      def scale(value, rawRange, scaledRange):
          def computeSlope(inputRange, outputRange):
              outputRangeDelta = outputRange[1] - outputRange[0]
              inputRangeDelta = inputRange[1] - inputRange[0]

              if (inputRangeDelta == 0):
                  return 0
              else:
                  return outputRangeDelta / inputRangeDelta
              end
          end

          def computeIntercept(slope, inputRange, outputRange):
              return outputRange[0] - (slope * inputRange[0])
          end

          def clipScaledValue(outputScaledValue, outputRange):
              if (outputRange[0] < outputRange[1]):
                  return clipWhenLowerLimitIsLessThanHigher(outputScaledValue, outputRange)
              else:
                  return clipWhenLowerLimitIsGreaterThanHigherLimit(outputScaledValue, outputRange)
              end
          end

          def clipWhenLowerLimitIsGreaterThanHigherLimit(outputScaledValue, outputRange):
              if (outputScaledValue < outputRange[1]):
                  return outputRange[1]
              elif (outputScaledValue > outputRange[0]):
                  return outputRange[0]
              else:
                  return outputScaledValue
              end
          end

          def clipWhenLowerLimitIsLessThanHigher(outputScaledValue, outputRange):
              if (outputScaledValue < outputRange[0]):
                  return outputRange[0]
              elif (outputScaledValue > outputRange[1]):
                  return outputRange[1]
              else:
                  return outputScaledValue
              end
          end

          slope = computeSlope(rawRange, scaledRange)
          intercept = computeIntercept(slope, rawRange, scaledRange)
          scaledValue = slope * value + intercept
          return clipScaledValue(scaledValue, scaledRange)
      end

      def limit(value, range):
          return scale(value, range, range)
      end


  rq_init_comm_if_connected(9, "1")
  rq_init_comm_if_connected(2, "2")
  rq_init_comm_if_connected(3, "3")
  rq_init_comm_if_connected(4, "4")
  rq_print_connected_grippers()
  rq_gripper_communication_thread = run rq_gripper_communication()
  set_closed_norm(97.6470588235294, "1")
  set_open_norm(1.1764705882352942, "1")
  set_closed_mm(0.0, "1")
  set_open_mm(53.0, "1")
  set_closed_norm(100.0, "2")
  set_open_norm(0.0, "2")
  set_closed_mm(0.0, "2")
  set_open_mm(50.0, "2")
  set_closed_norm(100.0, "3")
  set_open_norm(0.0, "3")
  set_closed_mm(0.0, "3")
  set_open_mm(50.0, "3")
  set_closed_norm(100.0, "4")
  set_open_norm(0.0, "4")
  set_closed_mm(0.0, "4")
  set_open_mm(50.0, "4")
  rq_current_limit_enabled = False
  while(not rq_gripper_communication_thread_started):
      sleep(0.008)
  end
  # end: URCap Installation Node
  step_count_300fee78_b3e2_4ecc_acea_62356c60d52b = 0.0
  thread Step_Counter_Thread_351342f9_30f5_4523_8313_4ca12f4a91f7():
    while (True):
      step_count_300fee78_b3e2_4ecc_acea_62356c60d52b = step_count_300fee78_b3e2_4ecc_acea_62356c60d52b + 1.0
      sync()
    end
  end
  run Step_Counter_Thread_351342f9_30f5_4523_8313_4ca12f4a91f7()
  global AMR_Position=struct(position_identifier=0, x1=0, x2=0, y1=0, y2=0, theta1=0, theta2=0)
  global CAM_Pose=p[0,0,0,0,0,0]
  global CAM_Relation=""
  global CMD_Abort=  False
  global CMD_Clear=  False
  global CMD_Reset=  False
  global CMD_Start=  False
  global CMD_Suspend=  False
  global CMD_Unhold=  False
  global CMD_Unsuspend=  False
  global CNT_Rack_Output=0
  global FNC_Freedrive=  False
  global PRC_TubCounter=0
  global STP=0
  global easyPickCount_4=0
  global easyPickCount_7=0
  global easyPickNoObj_4=0
  global easyPickNoObj_7=0
  global easyPickParts_4=0
  global easyPickParts_7=0
  global TMR_Barcode=0
  global Container_mid_1_p=p[-.379239199143, -.127191311915, .299999999998, .000000000046, -.000000000021, -1.247199999994]
  global Container_mid_1_q=[-2.477408934449926, -1.2969853503591224, -1.875639182904262, -1.539621866126728, 1.5731943360401213, -2.8009955944022717]
  global trigger_otw_p=p[-.364831738276, -.163967193938, .343299997821, .000000000046, -.000000000020, -1.148401333327]
  global trigger_otw_q=[-2.378283213085033, -1.2994862387706814, -1.7634300687554951, -1.6493302004167063, 1.573123683454141, -2.8011223671816943]
  global Waypoint_54_p=p[.008800512419, -.547926542621, .402696567415, -.589884378425, -.007228654778, -.061268144704]
  global Waypoint_54_q=[-1.2044575850116175, -1.3416667741588135, -1.8272563219070435, -0.9884541195682068, 1.3621035814285278, -2.7712565104113978]
  global Waypoint_77_p=p[-.178371829612, -.433927395311, .368082383916, -.086593488055, .704679941724, -.007869906074]
  global Waypoint_77_q=[-1.265390698109762, -1.3355963987163086, -1.7944865226745605, -1.7402602634825648, 0.8780410885810852, -2.7713127771960657]
  global Waypoint_83_p=p[.008800512419, -.547926542621, .402696567415, -.589884378425, -.007228654778, -.061268144704]
  global Waypoint_83_q=[-1.2044575850116175, -1.3416667741588135, -1.8272563219070435, -0.9884541195682068, 1.3621035814285278, -2.7712565104113978]
  global Waypoint_84_p=p[-.178371829612, -.433927395311, .368082383916, -.086593488055, .704679941724, -.007869906074]
  global Waypoint_84_q=[-1.265390698109762, -1.3355963987163086, -1.7944865226745605, -1.7402602634825648, 0.8780410885810852, -2.7713127771960657]
  global Vial_above_1_p=p[.017105793010, -.652093028359, .184920586844, .000000000272, .000000000270, 1.564063451276]
  global Vial_above_1_q=[-1.3375440709712851, -1.9618096977868804, -1.4665759083780685, -1.2837941559171444, 1.5732503672317195, -4.47276330421513]
  global Vial_pick_poi_1_p=p[.017105792852, -.648922724010, .093307568731, .000000000271, .000000000270, 1.564063451276]
  global Vial_pick_poi_1_q=[-1.3366329456391917, -2.0375277831965413, -1.6071432798879028, -1.0675084332049813, 1.57309887265915, -4.471135348858068]
  global Waypoint_86_p=p[.019227646885, -.648669633640, .184920586950, .000000000000, .000000000000, .024063451426]
  global Waypoint_86_q=[-1.3331129109407733, -1.9540750545686123, -1.4775914902901128, -1.280581784992414, 1.5733500744865856, -2.928303704452631]
  global Waypoint_87_p=p[-.032361834699, -.348336136197, .391475576335, -.000008499254, .000014589902, -.004651426820]
  global Waypoint_87_q=[-1.2709335019096129, -1.1914598663441005, -1.708995335060501, -1.8117888533498316, 1.5729683532263925, -2.8379347397710237]
  global Vial_3FG_plac_1_p=p[-.031858676359, -.349402499566, .145301120695, .000000000000, .000000000000, .000000000000]
  global Vial_3FG_plac_1_q=[-1.2723975525801707, -1.252376585823825, -2.3128114007049496, -1.1470592278900167, 1.5730548099411423, -2.8414815174610535]
  global Waypoint_88_p=p[-.032361834699, -.348336136197, .391475576335, -.000008499254, .000014589902, -.004651426820]
  global Waypoint_88_q=[-1.2709335019096129, -1.1914598663441005, -1.708995335060501, -1.8117888533498316, 1.5729683532263925, -2.8379347397710237]
  global cap_dump_1_p=p[-.139168676487, -.420163541420, .146096395183, .000000000000, .000000000000, .000000000000]
  global cap_dump_1_q=[-1.584588644510994, -1.5093464179777323, -2.1118449369620347, -1.091059703602438, 1.5728943834877336, -3.154014906686923]
  global Waypoint_89_p=p[-.032361834699, -.348336136197, .391475576335, -.000008499254, .000014589902, -.004651426820]
  global Waypoint_89_q=[-1.2709335019096129, -1.1914598663441005, -1.708995335060501, -1.8117888533498316, 1.5729683532263925, -2.8379347397710237]
  global Vial_3FG_plac_2_p=p[-.031858676359, -.349402499566, .145301120695, .000000000000, .000000000000, .000000000000]
  global Vial_3FG_plac_2_q=[-1.2723975525801707, -1.252376585823825, -2.3128114007049496, -1.1470592278900167, 1.5730548099411423, -2.8414815174610535]
  global Waypoint_90_p=p[-.032361834699, -.348336136197, .391475576335, -.000008499254, .000014589902, -.004651426820]
  global Waypoint_90_q=[-1.2709335019096129, -1.1914598663441005, -1.708995335060501, -1.8117888533498316, 1.5729683532263925, -2.8379347397710237]
  global cap_dump_2_p=p[-.139168676487, -.420163541420, .146096395183, .000000000000, .000000000000, .000000000000]
  global cap_dump_2_q=[-1.584588644510994, -1.5093464179777323, -2.1118449369620347, -1.091059703602438, 1.5728943834877336, -3.154014906686923]
  global Waypoint_91_p=p[-.032361834699, -.348336136197, .391475576335, -.000008499254, .000014589902, -.004651426820]
  global Waypoint_91_q=[-1.2709335019096129, -1.1914598663441005, -1.708995335060501, -1.8117888533498316, 1.5729683532263925, -2.8379347397710237]
  global Vial_liq_abov_1_p=p[-.025303660977, -.338758622354, .426628485936, -1.315858642253, .800043520260, -.928295855026]
  global Vial_liq_abov_1_q=[-0.3789628187762659, -1.5149522957256814, -2.263045310974121, 0.7870649534412841, -0.750984017048971, -3.2237566153155726]
  global Vial_liq_pick_3_p=p[-.002660428945, -.335984893034, .159389832934, -1.150456778400, .673175527684, -1.010612657503]
  global Vial_liq_pick_3_q=[-0.3660772482501429, -1.4503649038127442, -2.4056053161621094, -1.994692941705221, 0.8039668202400208, -0.2508929411517542]
  global Vial_liq_pick_4_p=p[-.041402486291, -.356791603314, .125395323246, -1.143483969075, .651070210027, -.878721885453]
  global Vial_liq_pick_4_q=[-0.4426233705502476, -1.437252121513727, -2.551930962114307, -1.776528229806984, 0.6562026234073748, -0.43018811960029524]
  global Vial_liq_abov_2_p=p[-.025303660977, -.338758622354, .426628485936, -1.315858642253, .800043520260, -.928295855026]
  global Vial_liq_abov_2_q=[-0.3789628187762659, -1.5149522957256814, -2.263045310974121, 0.7870649534412841, -0.750984017048971, -3.2237566153155726]
  global Liquid_midway_1_p=p[.057575295009, -.583081747994, .306414980749, -1.351675548728, .120935756539, -.096908606303]
  global Liquid_midway_1_q=[-0.895174805318014, -1.7035466633238734, -2.380953073501587, 0.631549521083496, 0.7706599235534668, -2.9455552736865442]
  global shake_3_p=p[.057574880217, -.583085370269, .306422893466, -1.360996190983, -.155555042453, -.438136255921]
  global shake_3_q=[-0.8951800505267542, -1.7035466633238734, -2.380937099456787, 0.6315542894550782, 0.7706599235534669, -2.5394540616517496]
  global shake_4_p=p[.057581636113, -.583090570002, .306439684073, -1.308767904323, .368530312677, .214926493520]
  global shake_4_q=[-0.8951714674579065, -1.7035395107665003, -2.380906343460083, 0.6315504747578125, 0.7706480026245118, -3.3161255787892268]
  global drop_above_3_p=p[.268235025993, -.467784390499, .226219872376, -1.027832627524, -.430841408251, 1.004603115937]
  global drop_above_3_q=[-0.935645882283346, -1.6663371525206507, -2.4252893924713135, 0.41966931402172847, 1.8470635414123535, -3.4600217978106897]
  global drop_above_4_p=p[.219042229014, -.470775657081, .133754190740, -.313004595901, -.344395319364, 1.500564994056]
  global drop_above_4_q=[-1.0601594887284795, -1.70046459045642, -2.0799996233759863, -0.7243227230676759, 1.9429634314685202, -4.115129153870795]
  global liq_tran_3_p=p[.213067510942, -.469567035397, .100231043184, .251862243732, .217902579404, 1.592812335393]
  global liq_tran_3_q=[-0.7789645168037476, -1.822364827406652, -1.8643518410805573, -1.252158963840138, 1.3768134449520435, -3.9328333233290254]
  global drop_above_5_p=p[.219042229014, -.470775657081, .133754190740, -.313004595901, -.344395319364, 1.500564994056]
  global drop_above_5_q=[-1.0601594887284795, -1.70046459045642, -2.0799996233759863, -0.7243227230676759, 1.9429634314685202, -4.115129153870795]
  global Waypoint_92_p=p[.187119460405, -.493959476151, .133754190608, -.313004596540, -.344395317757, 1.500564993991]
  global Waypoint_92_q=[-1.1418328121400876, -1.7310553375189475, -2.033634768766424, -0.772026910513711, 1.958578934631971, -4.201588449364511]
  global liq_tran_4_p=p[.195957706507, -.493022614126, .100231042689, .160718757180, .109807038912, 1.525321508623]
  global liq_tran_4_q=[-0.881740380645474, -1.8244526267589851, -1.865100964490387, -1.1608866323693583, 1.4631433601076713, -3.973915130363038]
  global drop_above_6_p=p[.219042229014, -.470775657081, .133754190740, -.313004595901, -.344395319364, 1.500564994056]
  global drop_above_6_q=[-1.0601594887284795, -1.70046459045642, -2.0799996233759863, -0.7243227230676759, 1.9429634314685202, -4.115129153870795]
  global drop_above_7_p=p[.268235025993, -.467784390499, .226219872376, -1.027832627524, -.430841408251, 1.004603115937]
  global drop_above_7_q=[-0.935645882283346, -1.6663371525206507, -2.4252893924713135, 0.41966931402172847, 1.8470635414123535, -3.4600217978106897]
  global Liquid_midway_2_p=p[.057575295009, -.583081747994, .306414980749, -1.351675548728, .120935756539, -.096908606303]
  global Liquid_midway_2_q=[-0.895174805318014, -1.7035466633238734, -2.380953073501587, 0.631549521083496, 0.7706599235534668, -2.9455552736865442]
  global Vial_drop_abo_1_p=p[.000324902251, -.648569523142, .221894115667, -.873462921366, 1.165852672573, -1.482720593185]
  global Vial_drop_abo_1_q=[-1.0576906334721352, -2.393016994184633, -0.9236232851859159, -2.5729213042279273, 0.7903331288549689, -0.33286325848155585]
  global Vial_liq_drop_1_p=p[.001020867953, -.647659915585, .092915870838, -.834762611599, 1.081942994823, -1.540647900176]
  global Vial_liq_drop_1_q=[-1.0631954168193474, -2.4447642951220825, -1.128811017825127, -2.1983115491972294, 0.8130148661460634, -0.38984988696911316]
  global Vial_drop_abo_2_p=p[.000324902251, -.648569523142, .221894115667, -.873462921366, 1.165852672573, -1.482720593185]
  global Vial_drop_abo_2_q=[-1.0576906334721352, -2.393016994184633, -0.9236232851859159, -2.5729213042279273, 0.7903331288549689, -0.33286325848155585]
  global Spatula_otw_p=p[-.038472058237, -.263141484147, .425351216717, -.000441582511, -.000128175490, 3.034387645854]
  global Spatula_otw_q=[-1.1888947506684495, -1.0083288774886814, -1.7052227056065874, -1.9984805067363443, 1.5730180972985317, 0.48793409320312264]
  global pick_spat_L_abv_p=p[.239059466375, -.067212518441, .280720723617, .000017217488, -.000484427718, 3.106837214660]
  global pick_spat_L_abv_q=[0.292765616142962, -0.8565557553273315, -2.140199892763044, -1.715349495646084, 1.573623142106424, 1.8984976776985687]
  global spat_L_pick_p=p[.242468789885, -.067301915011, .193171208067, .000017217488, -.000484427718, 3.106837214657]
  global spat_L_pick_q=[0.2867414378807389, -0.8600077002089179, -2.3629148016312627, -1.4891831672860159, 1.5737695566221115, 1.8933890858591198]
  global spat_L_lift_p=p[.245402002494, -.067432373551, .289049296496, .000017217490, -.000484427724, 3.106837214657]
  global spat_L_lift_q=[0.2834351187564135, -0.8798320076811592, -2.1119436738532986, -1.7203314352121302, 1.573588313403067, 1.8891054681654005]
  global spat_L_side_p=p[.247133573905, -.017633681797, .289062935631, .000017217490, -.000484427724, 3.106837214657]
  global spat_L_side_q=[0.49719173575848863, -0.8582398211168538, -2.1182130454788215, -1.735610316654931, 1.5735817737572706, 2.1028402698705397]
  global spat_L_up_p=p[.247135508752, -.017665230822, .397130746165, .000017217490, -.000484427724, 3.106837214657]
  global spat_L_up_q=[0.49854946074076967, -0.9346239623559676, -1.808280269374471, -1.969158816463132, 1.5731020084036995, 2.1031742024348157]
  global spat_M_up_p=p[.245495561680, -.112112573515, .420343789747, .000026293989, -.000477463067, 3.067686800858]
  global spat_M_up_q=[0.09017908059107435, -1.0134242235449396, -1.71728844067247, -1.9814399845077446, 1.573013686840385, 1.733759055129931]
  global spat_M_pick_p=p[.244673518506, -.111985070134, .192299022723, .000026293990, -.000477463072, 3.067686800901]
  global spat_M_pick_q=[0.08834054082534859, -0.9272467647495475, -2.3438023910348154, -1.4411029496965373, 1.5736983399628084, 1.7342144371718433]
  global spat_S_Up_7_p=p[.252087445596, -.159242094834, .423281604617, .000026293954, -.000477463070, 3.067686800855]
  global spat_S_Up_7_q=[-0.09804692328730358, -1.0862987822056382, -1.6788706463996483, -1.9470242450550348, 1.5730147401359813, 1.5455107082823842]
  global spat_S_Pick_4_p=p[.245377020686, -.158668022535, .192285730279, .000026293985, -.000477463062, 3.067686800840]
  global spat_S_Pick_4_q=[-0.10087203759495189, -1.011188488703386, -2.311978084495874, -1.3890267520590838, 1.5735990551056096, 1.5450562970948172]
  global spat_S_Up_8_p=p[.252087445596, -.159242094834, .423281604617, .000026293954, -.000477463070, 3.067686800855]
  global spat_S_Up_8_q=[-0.09804692328730358, -1.0862987822056382, -1.6788706463996483, -1.9470242450550348, 1.5730147401359813, 1.5455107082823842]
  global spat_flatM_up_p=p[.229022666361, -.211442909333, .418634047126, .000026293953, -.000477463083, 3.067686800888]
  global spat_flatM_up_q=[-0.30183372580416545, -1.1157042924275036, -1.6775646144685776, -1.9189678841796578, 1.5730340557943228, 1.341766142011193]
  global spat_flatM_pick_p=p[.241028983327, -.208057297586, .192270533170, .000026293950, -.000477463079, 3.067686800885]
  global spat_flatM_pick_q=[-0.2805687960562633, -1.1003763929487214, -2.271431297337675, -1.3404236887924883, 1.5734924238720627, 1.3653813047742556]
  global spat_flatS_up_p=p[.237651953780, -.253943828614, .403961222825, .000026293950, -.000477463092, 3.067686800841]
  global spat_flatS_up_q=[-0.42363550926974103, -1.1939944599502539, -1.6745915127240307, -1.843675057902054, 1.5731001874678698, 1.220082820532415]
  global spat_flatS_pick_p=p[.241325662334, -.251726327528, .192256842740, .000026293947, -.000477463087, 3.067686800841]
  global spat_flatS_pick_q=[-0.4144907797170738, -1.1967447109013012, -2.21926362252748, -1.2962499335425761, 1.5733885098427622, 1.2314402238866728]
  global spat_S_pick_p=p[.238158866340, -.157926795425, .192632100345, .000026293989, -.000477463069, 3.067686800857]
  global spat_S_pick_q=[-0.10084756991493293, -0.9881392730064915, -2.3204232610157494, -1.403630829593915, 1.5736254260650586, 1.5450653591083503]
  global spat_S_up_p=p[.244260523725, -.164466690315, .417087579736, .000026293988, -.000477463072, 3.067686800857]
  global spat_S_up_q=[-0.12101499604198729, -1.0718307017854336, -1.7023391702814736, -1.938028805938881, 1.573044424728474, 1.5226045951991447]
  global Waypoint_7_p=p[-.472820924474, .292439826233, .207418370237, -.137787250486, 2.177332259632, -2.152029714756]
  global Waypoint_7_q=[-2.911134078210732, -1.90240864358569, -1.968768330510411, -2.500365101593811, 0.11427687110891149, 0.0958980389250167]
  global Waypoint_8_p=p[-.357612884176, -.251084817998, .212379799667, -.858181193174, 1.714832512191, -1.687547565568]
  global Waypoint_8_q=[-1.620834863369681, -1.8936194567376496, -1.9821394403832038, -2.4599791457905273, 0.6296693672615152, 0.07625365420707819]
  global Decapp_above_3_p=p[-.013480295948, -.359153355979, .266194408367, -.879653555922, 1.646336924805, -1.709111068605]
  global Decapp_above_3_q=[-0.9632157249872035, -2.0163405763031657, -1.5968194594157152, -2.6579215719847085, 1.251243398585566, 0.047906446502667066]
  global Decapp_place_3_p=p[-.013480295890, -.359153356055, .160907502384, -.879653554902, 1.646336919740, -1.709111066456]
  global Decapp_place_3_q=[-0.9633402410919709, -2.1541179572356635, -1.6937729380888573, -2.4232786481058053, 1.2517342187662468, 0.04818402956922263]
  global Decapp_above_4_p=p[-.013480295948, -.359153355979, .266194408367, -.879653555922, 1.646336924805, -1.709111068605]
  global Decapp_above_4_q=[-0.9632157249872035, -2.0163405763031657, -1.5968194594157152, -2.6579215719847085, 1.251243398585566, 0.047906446502667066]
  global Waypoint_78_p=p[-.051450028091, -.519555688329, .365718563414, -1.287302938145, 1.077637394477, -1.218524965834]
  global Waypoint_78_q=[-0.9214276262416012, -1.8899696965062578, -1.4939326452510562, -2.840015661555725, 0.5585157189668353, 0.033997638875617575]
  global Waypoint_10_p=p[-.330595116596, .282932669854, .220236276291, 1.304675539882, .014233792938, -1.753932442581]
  global Waypoint_10_q=[-3.189526379253601, -1.8418198435143305, -1.7138504750370807, -2.182789974066381, 1.0126080912871243, -2.4455984844694645]
  global Waypoint_9_p=p[-.538777454962, .370695704977, .175030018143, -.317104215445, 2.082346543003, -2.037631421082]
  global Waypoint_9_q=[-3.1158871966457857, -1.998548595120492, -1.941797010061462, -2.2703530575838844, -0.27573365931009164, -0.06926782177267654]
  global Powder_wayp1_p=p[-.472820924474, .292439826233, .207418370237, -.137787250486, 2.177332259632, -2.152029714756]
  global Powder_wayp1_q=[-2.911134078210732, -1.90240864358569, -1.968768330510411, -2.500365101593811, 0.11427687110891149, 0.0958980389250167]
  global Waypoint_2_p=p[-.357612884176, -.251084817998, .212379799667, -.858181193174, 1.714832512191, -1.687547565568]
  global Waypoint_2_q=[-1.620834863369681, -1.8936194567376496, -1.9821394403832038, -2.4599791457905273, 0.6296693672615152, 0.07625365420707819]
  global Postions_otw_p=p[-.010896578244, -.533368729951, .288851175116, -1.233738470894, 1.195331112012, -1.207314088469]
  global Postions_otw_q=[-0.898791023514228, -2.078490033037677, -1.4499891355755317, -2.7624416226992476, 0.6570218891920963, 0.02136606178275929]
  global cont_A_otw_p=p[.070238108556, -.655257851554, .184611566008, -1.090601381517, 1.404822685081, -1.413645380264]
  global cont_A_otw_q=[-0.990969136335913, -2.7123780097559784, -0.5772671651193146, -3.0005537851220403, 0.84719335943793, 0.020652463706785973]
  global cont_B_otw_p=p[.256012899886, -.515433666916, .157862612232, -1.209199576153, 1.209199576154, -1.209199576153]
  global cont_B_otw_q=[-0.6068713783523112, -2.5251567701153963, -1.0126698074772102, -2.742679391438185, 0.9631140738765777, -0.0042246938882417595]
  global cont_C_otw_p=p[.319495487998, -.362719410364, .163846736977, -1.233784872294, 1.195277203291, -1.207325031551]
  global cont_C_otw_q=[-0.3611889651645974, -2.404603865546651, -1.2341573845076566, -2.650535279811077, 1.1944844573128257, 0.01638086594640864]
  global Waypoint_1_p=p[-.352029261722, -.424157832422, .472326578019, -.000004407962, .000020663369, -1.529709227737]
  global Waypoint_1_q=[-2.017015745614491, -1.7423968528991196, -1.0053357238485425, -1.9644715035904907, 1.5727249689896, -2.060727852912713]
  global Waypoint_5_p=p[.219993437017, -.447144142811, .462350040687, .000006087494, .000031090075, .000022232405]
  global Waypoint_5_q=[-0.8406239476037944, -1.5982534362206806, -1.1934200873248484, -1.9205794898315975, 1.5727336676986443, -2.4135960466995314]
  global cont_B_safe_p=p[.256012900841, -.515433666823, .234963258529, -1.209199574203, 1.209199576702, -1.209199577238]
  global cont_B_safe_q=[-0.5984778117169087, -2.477204487479997, -0.8976875250023646, -2.905631546928806, 0.9709012567976698, -0.00424039942746024]
  global PosA_up_p=p[.028578953747, -.638006009765, .227275735849, -1.090660933958, 1.404791542934, -1.413645191233]
  global PosA_up_q=[-1.0254743496427432, -2.565176838504783, -0.7558042274983681, -2.9696064674274343, 0.8129191411995651, 0.021444818458024387]
  global PosA_pick_p=p[.026918718687, -.640084889741, .097901147521, -1.090660933959, 1.404791542934, -1.413645191233]
  global PosA_pick_q=[-1.028821435558534, -2.6899890636403807, -0.8526126047665157, -2.7478942693937167, 0.8103607002888742, 0.021326778146411485]
  global PosB_up_p=p[.239472634782, -.492481416782, .220767759213, -1.233738470883, 1.195331111998, -1.207314088469]
  global PosB_up_q=[-0.5800230603397054, -2.4076296700885997, -1.0699783327330836, -2.8116344407747427, 0.9750472858169287, 0.017627507888886562]
  global PosB_pick_p=p[.240630296955, -.494558620171, .096392895280, -1.233740573549, 1.195309876041, -1.207293779132]
  global PosB_pick_q=[-0.5816146260408139, -2.553273721769836, -1.1376320925804277, -2.5983292591462153, 0.9740936784345416, 0.017625262979849232]
  global PosC_up_p=p[.241566602786, -.359249123455, .230260583862, -1.233738470888, 1.195331111997, -1.207314088449]
  global PosC_up_q=[-0.39573787962534546, -2.2019009616581497, -1.4115270142506517, -2.675987785326166, 1.160180741930842, 0.01687917643039505]
  global PosC_pick_p=p[.240633854030, -.361553124916, .093979792658, -1.233738470878, 1.195331111997, -1.207314088469]
  global PosC_pick_q=[-0.39992427526118757, -2.386042391328985, -1.4894374567278712, -2.414022930893381, 1.1566786195951169, 0.01712017454263659]
  global Pow_decap_up_p=p[-.017556487132, -.367519866742, .275835445416, -.605635182849, 1.892518157522, -1.890848751165]
  global Pow_decap_up_q=[-1.1272088681128203, -2.1173924123331025, -1.4250048354055203, -2.7485980486387676, 1.4193896902217862, 0.023247957637719453]
  global pow_decap_place_p=p[-.020433194420, -.368310202914, .161281291611, -.605635182838, 1.892518157522, -1.890848751163]
  global pow_decap_place_q=[-1.132360890531647, -2.2521863255983092, -1.5302136899970318, -2.5086176644751683, 1.4149282844269635, 0.02347140074572661]
  global Decap_above_p=p[-.031863883354, -.349974838955, .288042264213, .000000000000, .000000000000, .000000000000]
  global Decap_above_q=[-1.271900116540503, -1.1670201114602632, -1.989291655468758, -1.5559360538518163, 1.573255119759632, -2.842476569674073]
  global Decapp_p=p[-.031864263150, -.349974612700, .230259377740, .000000000000, .000000000000, .000000000000]
  global Decapp_q=[-1.2723555431601419, -1.1810456878410935, -2.1291754890757737, -1.4020263844320349, 1.5732701843074919, -2.842325632263757]
  global Cap_above_p=p[-.224192409203, -.629599568633, .257274081142, .000015605575, -.000015166009, -1.647823825902]
  global Cap_above_q=[-1.710642681834492, -1.9674285251810462, -1.2705185053146897, -1.4742193161331247, 1.573506065067499, -1.6347709465008595]
  global Cap_place_p=p[-.224189049846, -.629597879697, .041885651757, .000015605572, -.000015166011, -1.647823825903]
  global Cap_place_q=[-1.7111696563854295, -2.13979870939016, -1.5941008764912503, -0.978265561728648, 1.5732789016410962, -1.6336328794662904]
  global OP_PowderA2_p=p[.009371277507, -.409434369247, .294169017766, -.823281033205, 1.709410851243, -1.698303593897]
  global OP_PowderA2_q=[-0.9994544761745754, -2.1395254572673217, -1.3437567783153916, -2.8143375616690456, 1.2617899549595724, 0.019614613715634555]
  global Decap_up_p=p[-.018339217391, -.367674469480, .249553854268, -.546164737599, 1.935964719000, -1.930057109666]
  global Decap_up_q=[-1.158124747223252, -2.1569920012936787, -1.4340832185069745, -2.7006032680036753, 1.4556626828962336, 0.02060977878679182]
  global Decap_pick_p=p[-.020429098827, -.367971872627, .161604333799, -.546164737600, 1.935964719000, -1.930057109666]
  global Decap_pick_q=[-1.161653098289774, -2.263509236689538, -1.5087211318402236, -2.519459740767391, 1.452646640403743, 0.02077912034002202]
  global Op_PowA_wP_p=p[-.173727579245, -.372934016396, .295116627479, -.972390492433, 1.540962074418, -1.548745344994]
  global Op_PowA_wP_q=[-1.1740587397768483, -1.865656321049359, -1.7426943793777419, -2.679427276872525, 0.8588908769087338, 0.017944699631825187]
  global TMR_Barcode_is_counting=False
  thread Timer_Thread():
    while (True):
      if (TMR_Barcode_is_counting):
        TMR_Barcode = TMR_Barcode + get_steptime()
      end
      sync()
    end
  end
  run Timer_Thread()
  def Sub_Vision_V18():
    $ 816 "Sub_Vision_V18" "noBreak"
    $ 817 "PreSettings"
    $ 818 "CAM_LM_Detected≔ False "
    global CAM_LM_Detected=  False
    $ 819 "CAM_Captures≔0"
    global CAM_Captures=0
    $ 820 "CAM_Pose≔p[0,0,0,0,0,0]"
    global CAM_Pose=p[0,0,0,0,0,0]
    $ 821 "CAM_LM_Refinmnt≔ False "
    global CAM_LM_Refinmnt=  False
    $ 822 "CAM_LM_Refined≔ False "
    global CAM_LM_Refined=  False
    $ 823 "CAM_LM_Deviatn≔p[0,0,0,0,0,0]"
    global CAM_LM_Deviatn=p[0,0,0,0,0,0]
    $ 824 "CAM_LM_ID≔0"
    global CAM_LM_ID=0
    $ 825 "CAM_Done≔ False "
    global CAM_Done=  False
    $ 826 "CAM_CNT_Obj≔0"
    global CAM_CNT_Obj=0
    $ 827 "CAM_Result = []"
    CAM_Result = []
    $ 828 "OBJ_Detected≔ False "
    global OBJ_Detected=  False
    $ 829 "FRM_Reference≔p[0,0,0,0,0,0]"
    global FRM_Reference=p[0,0,0,0,0,0]
    $ 830 "'=========='"
    # '=========='
    $ 831 "Switch Action"
    switch_1 = Action
    $ 832 "Case 13"
    if (13 == switch_1):
    elif (15 == switch_1):
      $ 950 "Case 15"
    elif (131 == switch_1):
      $ 996 "Case 131"
      $ 997 "Read (SensoPart)"
      $ 998 "Action_Info≔'search for landmark'"
      global Action_Info="search for landmark"
      $ 999 "CAM_LM≔CAM_LMs[4]"
      global CAM_LM=CAM_LMs[4]
      $ 1000 "CAM_Relation≔CAM_LM.capture_relation"
      global CAM_Relation=CAM_LM.capture_relation
      $ 1001 "go to capture pose"
      $ 1004 "If ITM_ID≟1 and JIG≟7"
      if (ITM_ID == 1  and  JIG == 7):
        $ 1005 "PSE_T≔uLM_Cap_SSRack"
        global PSE_T=uLM_Cap_SSRack
      else:
        $ 1006 "ElseIf ITM_ID≟5 and JIG≟7"
        if (ITM_ID == 5  and  JIG == 7):
          $ 1007 "PSE_T≔FRM_Cap_SSRack"
          global PSE_T=FRM_Cap_SSRack
        else:
          $ 1010 "ElseIf ITM_ID≟1 and JIG≟15"
          if (ITM_ID == 1 and JIG == 15):
            $ 1011 "MoveJ"
            $ 1012 "Container_mid_1" "breakAfter"
            movej(get_inverse_kin(Container_mid_1_p, qnear=Container_mid_1_q), a=1.3962634015954636, v=1.0471975511965976, r=0.05)
            $ 1014 "PSE_T≔FRM_Container_const"
            global PSE_T=p[-0.5003348223692186,0.35061804815168285,0.41579001388808423,-5.092943187272062E-5,1.0145185065363121E-4,-2.764319258713288]
          else:
            $ 1015 "ElseIf ITM_ID≟1 and JIG≟21"
            if (ITM_ID == 1 and JIG == 21):
              $ 1016 "PSE_T≔FRM_PoTS_const"
              global PSE_T=p[-0.5403054403210852,-0.10910773999775857,0.4828,3.058497512721046E-6,2.3454853329357316E-5,-2.208510541952706]
            else:
              $ 1017 "ElseIf ITM_ID≟1 and JIG≟17"
              if (ITM_ID == 1 and JIG == 17):
                $ 1018 "MoveJ"
                $ 1019 "trigger_otw" "breakAfter"
                movej(get_inverse_kin(trigger_otw_p, qnear=trigger_otw_q), a=1.3962634015954636, v=1.0471975511965976, r=0.05)
                $ 1023 "PSE_T≔FRM_weigh_scale_const"
                global PSE_T=p[-0.3804866881697204,0.025744252835212,0.4723487455232425,-1.0445769542396123E-4,-1.924788411074358E-5,-2.1691978730572363]
              end
            end
          end
        end
      end
      $ 1024 "do_transition(PSE_T, keep_rxry=False)"
      do_transition(PSE_T, keep_rxry=False)
      $ 1025 "Set"
      set_tcp(p[0.0,0.0,0.161,3.1415,0.0,0.0])
      $ 1026 "MoveJ"
      $ 1027 "PSE_T" "breakAfter"
      movej(PSE_T, a=1.3962634015954636, v=1.7453292519943295)
      $ 1028 "CAM_Pose≔get_actual_tcp_pose()"
      global CAM_Pose= get_actual_tcp_pose ()
      $ 1029 "Loop  not CAM_Done and  not ERROR.FLAG and  not CMD_Stop"
      while (  not  CAM_Done  and    not  ERROR.FLAG  and    not  CMD_Stop):
        $ 1030 "adjust capture pose"
        $ 1031 "If CAM_LM_Detected and CAM_LM_Refinmnt"
        if (CAM_LM_Detected  and  CAM_LM_Refinmnt):
          $ 1032 "PSE_T≔p[0,0,0.300,0,0,0]"
          global PSE_T=p[0,0,0.300,0,0,0]
          $ 1033 "CAM_Pose≔PSE_T"
          global CAM_Pose=PSE_T
          $ 1034 "If  not is_reachable(FRM_Reference,[PSE_T])"
          if (  not  is_reachable(FRM_Reference,[PSE_T])):
            $ 1035 "Error"
            $ 1036 "set_error(ERROR_POSE_NOT_REACHABLE)"
            set_error(ERROR_POSE_NOT_REACHABLE)
          end
          $ 1037 "If  not ERROR.FLAG"
          if (  not  ERROR.FLAG):
            $ 1038 "MoveJ"
            $ 1039 "PSE_T" "breakAfter"
            set_tcp(p[0.0,0.0,0.161,0.0,0.0,0.0])
            movej(pose_trans(FRM_Reference, PSE_T), a=0.8726646259971648, v=1.3962634015954636)
            $ 1040 "CAM_LM_Refined≔ True "
            global CAM_LM_Refined=  True
          end
        else:
          $ 1041 "ElseIf  not CAM_LM_Detected and CAM_Captures>0"
          if (  not  CAM_LM_Detected  and  CAM_Captures>0):
            $ 1042 "MoveL"
            $ 1043 "If FRM_Reference≟p[0,0,0,0,0,0]"
            if (FRM_Reference == p[0,0,0,0,0,0]):
              $ 1044 "PSE_T≔get_random_pose(pose_ref=CAM_Pose, mode='cubic', range_max=[0.150,0.150,0.015])"
              global PSE_T=get_random_pose(pose_ref=CAM_Pose, mode="cubic", range_max=[0.150,0.150,0.015])
            else:
              $ 1049 "Else" "noBreak"
              $ 1050 "PSE_T≔get_random_pose(pose_ref=CAM_Pose, mode='rotation', range_max=[10,10,0])"
              global PSE_T=get_random_pose(pose_ref=CAM_Pose, mode="rotation", range_max=[10,10,0])
              $ 1051 "CAM_LM_Refined≔ True "
              global CAM_LM_Refined=  True
            end
            $ 1052 "If get_inverse_kin_has_solution(pose_trans(FRM_Reference, PSE_T))"
            if (get_inverse_kin_has_solution( pose_trans (FRM_Reference, PSE_T))):
              $ 1053 "Comment"
              # Comment
              $ 1054 "PSE_T" "breakAfter"
              set_tcp(p[0.0,0.0,0.161,3.1415,0.0,0.0])
              movel(pose_trans(FRM_Reference, PSE_T), a=0.03, v=0.05)
            else:
              $ 1055 "Else" "noBreak"
              $ 1056 "'If random pose is out of reach, set the initial cam pose'"
              # 'If random pose is out of reach, set the initial cam pose'
              $ 1057 "PSE_T≔CAM_Pose"
              global PSE_T=CAM_Pose
            end
          end
        end
        $ 1058 "Wait: 2.0"
        sleep(2.0)
        $ 1059 "trigger"
        $ 1060 "If ITM_ID≟1 and JIG≟7"
        if (ITM_ID == 1  and  JIG == 7):
          # begin: URCap Program Node
          #   Source: SensoPart VISOR Robotic, 2.0.6, SensoPart Industriesensorik GmbH
          #   Type: VISOR Trigger
          $ 1061 "# 1 VISOR Trigger"
          visor_changeJob(1, "Landmark_INVITE_2", 6000)
          visor_trigger(1, 6000, "arm")
          # end: URCap Program Node
        else:
          $ 1062 "ElseIf ITM_ID≟5 and JIG≟7"
          if (ITM_ID == 5  and  JIG == 7):
            # begin: URCap Program Node
            #   Source: SensoPart VISOR Robotic, 2.0.6, SensoPart Industriesensorik GmbH
            #   Type: VISOR Trigger
            $ 1063 "# 1 VISOR Trigger"
            visor_changeJob(1, "Landmark_INVITE_2", 6000)
            visor_trigger(1, 6000, "arm")
            # end: URCap Program Node
          else:
            $ 1064 "ElseIf ITM_ID≟13 and JIG≟7"
            if (ITM_ID == 13  and  JIG == 7):
              # begin: URCap Program Node
              #   Source: SensoPart VISOR Robotic, 2.0.6, SensoPart Industriesensorik GmbH
              #   Type: VISOR Trigger
              $ 1065 "# 1 VISOR Trigger"
              visor_changeJob(1, "Landmark_INVITE_2", 6000)
              visor_trigger(1, 6000, "arm")
              # end: URCap Program Node
            else:
              $ 1066 "ElseIf ITM_ID≟1 and JIG≟15"
              if (ITM_ID == 1 and JIG == 15):
                # begin: URCap Program Node
                #   Source: SensoPart VISOR Robotic, 2.0.6, SensoPart Industriesensorik GmbH
                #   Type: VISOR Trigger
                $ 1067 "# 1 VISOR Trigger"
                visor_changeJob(1, "Aztec_no_dot_pick", 6000)
                visor_trigger(1, 6000, "arm")
                # end: URCap Program Node
              else:
                $ 1068 "ElseIf ITM_ID≟1 and JIG≟21"
                if (ITM_ID == 1 and JIG == 21):
                  # begin: URCap Program Node
                  #   Source: SensoPart VISOR Robotic, 2.0.6, SensoPart Industriesensorik GmbH
                  #   Type: VISOR Trigger
                  $ 1069 "# 1 VISOR Trigger"
                  visor_changeJob(1, "PoTS", 6000)
                  visor_trigger(1, 6000, "arm")
                  # end: URCap Program Node
                else:
                  $ 1070 "ElseIf ITM_ID≟1 and JIG≟17"
                  if (ITM_ID == 1 and JIG == 17):
                    # begin: URCap Program Node
                    #   Source: SensoPart VISOR Robotic, 2.0.6, SensoPart Industriesensorik GmbH
                    #   Type: VISOR Trigger
                    $ 1071 "# 1 VISOR Trigger"
                    visor_changeJob(1, "Weigh_target", 6000)
                    visor_trigger(1, 6000, "arm")
                    # end: URCap Program Node
                  end
                end
              end
            end
          end
        end
        $ 1075 "TM_3D_Found≔visor_partsFound(1)"
        global TM_3D_Found= visor_partsFound (1)
        $ 1077 "If TM_3D_Found>0"
        if (TM_3D_Found>0):
          $ 1078 "CAM_LM_Detected≔ True "
          global CAM_LM_Detected=  True
          $ 1079 "CAM_Captures≔0"
          global CAM_Captures=0
        else:
          $ 1080 "Else" "noBreak"
          $ 1081 "CAM_LM_Detected≔ False "
          global CAM_LM_Detected=  False
          $ 1082 "CAM_Captures≔CAM_Captures+1"
          global CAM_Captures=CAM_Captures+1
        end
        $ 1087 "result"
        $ 1088 "If CAM_LM_Detected"
        if (CAM_LM_Detected):
          $ 1089 "If (CAM_LM_Refinmnt and CAM_LM_Refined) or  not CAM_LM_Refinmnt"
          if ((CAM_LM_Refinmnt  and  CAM_LM_Refined)  or    not  CAM_LM_Refinmnt):
            $ 1147 "If ITM_ID≟1 and JIG≟7"
            if (ITM_ID == 1  and  JIG == 7):
              $ 1148 "CAM_LM_SSRack≔visor_getPose3d(1, 0)"
              global CAM_LM_SSRack= visor_getPose3d (1, 0)
            else:
              $ 1149 "ElseIf ITM_ID≟5 and JIG≟7"
              if (ITM_ID == 5  and  JIG == 7):
                $ 1150 "CAM_LM_SSRack≔visor_getPose3d(1, 0)"
                global CAM_LM_SSRack= visor_getPose3d (1, 0)
              else:
                $ 1153 "ElseIf ITM_ID≟1 and JIG≟15"
                if (ITM_ID == 1 and JIG == 15):
                  $ 1154 "CAM_LM_cont≔visor_getPose3d(1, 0)"
                  global CAM_LM_cont= visor_getPose3d (1, 0)
                  $ 1155 "Trigger≔get_actual_tcp_pose()"
                  global Trigger= get_actual_tcp_pose ()
                else:
                  $ 1156 "ElseIf ITM_ID≟1 and JIG≟21"
                  if (ITM_ID == 1 and JIG == 21):
                    $ 1157 "CAM_LM_cont≔visor_getPose3d(1, 0)"
                    global CAM_LM_cont= visor_getPose3d (1, 0)
                    $ 1158 "Trigger≔get_actual_tcp_pose()"
                    global Trigger= get_actual_tcp_pose ()
                  else:
                    $ 1159 "ElseIf ITM_ID≟1 and JIG≟17"
                    if (ITM_ID == 1 and JIG == 17):
                      $ 1160 "CAM_LM_cont≔visor_getPose3d(1, 0)"
                      global CAM_LM_cont= visor_getPose3d (1, 0)
                      $ 1161 "Trigger≔get_actual_tcp_pose()"
                      global Trigger= get_actual_tcp_pose ()
                    end
                  end
                end
              end
            end
            $ 1162 "CAM_Done≔ True "
            global CAM_Done=  True
          end
        else:
          $ 1163 "ElseIf  not CAM_LM_Detected and CAM_Captures<CAM_PRM_Retries"
          if (  not  CAM_LM_Detected  and  CAM_Captures<CAM_PRM_Retries):
            $ 1164 "CAM_LM_Refined≔ False "
            global CAM_LM_Refined=  False
          else:
            $ 1165 "ElseIf CAM_Captures≥CAM_PRM_Retries"
            if (CAM_Captures >= CAM_PRM_Retries):
              $ 1166 "CAM_Done≔ True "
              global CAM_Done=  True
              $ 1167 "Error"
              $ 1168 "set_error(ERROR_NO_LANDMARK)"
              set_error(ERROR_NO_LANDMARK)
            end
          end
        end
      end
    elif (151 == switch_1):
      $ 1169 "Case 151"
      $ 1170 "Detect (SensoPart)"
      $ 1171 "go to capture pose"
      $ 1172 "FRM_Reference≔FRM_Cap_SSRack"
      global FRM_Reference=FRM_Cap_SSRack
      $ 1173 "PSE_T≔p[0,0,-0.00,0,0,0]"
      global PSE_T=p[0,0,-0.00,0,0,0]
      $ 1174 "do_transition(pose_trans(FRM_Reference, PSE_T), keep_rxry=False)"
      do_transition( pose_trans (FRM_Reference, PSE_T), keep_rxry=False)
      $ 1175 "JNT_Q≔get_actual_joint_positions()"
      global JNT_Q= get_actual_joint_positions ()
      $ 1176 "JNT_Q≔[JNT_Q[0], JNT_Q[1], JNT_Q[2], JNT_Q[3], JNT_Q[4], 0]"
      global JNT_Q=[JNT_Q[0], JNT_Q[1], JNT_Q[2], JNT_Q[3], JNT_Q[4], 0]
      $ 1177 "Set"
      set_tcp(p[0.0,0.0,0.161,3.1415,0.0,0.0])
      $ 1178 "movej(get_inverse_kin(pose_trans(FRM_Reference, PSE_T), qnear=JNT_Q))"
      movej(get_inverse_kin( pose_trans (FRM_Reference, PSE_T), qnear=JNT_Q))
      $ 1179 "CAM_Pose≔pose_trans(pose_inv(FRM_Reference), get_actual_tcp_pose())"
      global CAM_Pose= pose_trans ( pose_inv (FRM_Reference),  get_actual_tcp_pose ())
      $ 1180 "Loop  not CAM_Done and  not ERROR.FLAG and  not CMD_Stop"
      while (  not  CAM_Done  and    not  ERROR.FLAG  and    not  CMD_Stop):
        $ 1181 "If  not OBJ_Detected and CAM_Captures>0"
        if (  not  OBJ_Detected  and  CAM_Captures>0):
          $ 1182 "MoveL"
          $ 1183 "If FRM_Reference≟p[0,0,0,0,0,0]"
          if (FRM_Reference == p[0,0,0,0,0,0]):
            $ 1185 "PSE_T≔get_random_pose(pose_ref=CAM_Pose, mode='rotation', range_max=[15,15,0])"
            global PSE_T=get_random_pose(pose_ref=CAM_Pose, mode="rotation", range_max=[15,15,0])
          else:
            $ 1186 "Else" "noBreak"
            $ 1187 "PSE_T≔get_random_pose(pose_ref=CAM_Pose, mode='rotation', range_max=[10,10,0])"
            global PSE_T=get_random_pose(pose_ref=CAM_Pose, mode="rotation", range_max=[10,10,0])
          end
          $ 1188 "If get_inverse_kin_has_solution(pose_trans(FRM_Reference, PSE_T))"
          if (get_inverse_kin_has_solution( pose_trans (FRM_Reference, PSE_T))):
            $ 1189 "PSE_T" "breakAfter"
            set_tcp(p[0.0,0.0,0.161,3.1415,0.0,0.0])
            movel(pose_trans(FRM_Reference, PSE_T), a=0.03, v=0.05)
          else:
            $ 1190 "Else" "noBreak"
            $ 1191 "'If random pose is out of reach, set the initial cam pose'"
            # 'If random pose is out of reach, set the initial cam pose'
            $ 1192 "PSE_T≔CAM_Pose"
            global PSE_T=CAM_Pose
            $ 1193 "PSE_T" "breakAfter"
            set_tcp(p[0.0,0.0,0.161,3.1415,0.0,0.0])
            movel(pose_trans(FRM_Reference, PSE_T), a=0.03, v=0.05)
          end
        end
        $ 1194 "Wait: 0.5"
        sleep(0.5)
        $ 1195 "Set"
        set_tcp(p[0.0,0.0,0.161,3.1415,0.0,0.0])
        # begin: URCap Program Node
        #   Source: SensoPart VISOR Robotic, 2.0.6, SensoPart Industriesensorik GmbH
        #   Type: VISOR Trigger
        $ 1196 "# 1 VISOR Trigger"
        visor_changeJob(1, "Object Detection Single", 6000)
        visor_trigger(1, 6000, "arm")
        # end: URCap Program Node
        $ 1197 "If visor_isResponseOk(1)"
        if ( visor_isResponseOk (1)):
          $ 1198 "CAM_CNT_Obj≔visor_partsFound(1)"
          global CAM_CNT_Obj= visor_partsFound (1)
          $ 1199 "CAM_OBJ_Pose≔visor_getPose3d(1, 0)"
          global CAM_OBJ_Pose= visor_getPose3d (1, 0)
          $ 1200 "If CAM_CNT_Obj>0"
          if (CAM_CNT_Obj>0):
            $ 1201 "CAM_OBJ_Color≔visor_getAdditionalData(1, 0)"
            global CAM_OBJ_Color= visor_getAdditionalData (1, 0)
            $ 1202 "CAM_DetectScore≔to_num(visor_getAdditionalData(1, 1))/1000"
            global CAM_DetectScore=to_num( visor_getAdditionalData (1, 1))/1000
            $ 1203 "OBJ_Detected≔ True "
            global OBJ_Detected=  True
          end
        else:
          $ 1204 "Else" "noBreak"
          $ 1205 "CAM_Captures≔CAM_Captures+1"
          global CAM_Captures=CAM_Captures+1
        end
        $ 1206 "If OBJ_Detected"
        if (OBJ_Detected):
          $ 1207 "Get object data"
          $ 1208 "PRC_CntDetect≔0"
          global PRC_CntDetect=0
          $ 1209 "Loop PRC_CntDetect<CAM_CNT_Obj"
          while (PRC_CntDetect<CAM_CNT_Obj):
            $ 1210 "get object and jig number"
            $ 1211 "If ITM_ID≟1 and JIG≟7"
            if (ITM_ID == 1  and  JIG == 7):
              $ 1212 "FRM_Reference≔FRM_Cap_SSRack"
              global FRM_Reference=FRM_Cap_SSRack
            else:
              $ 1213 "ElseIf ITM_ID≟5 and JIG≟7"
              if (ITM_ID == 5  and  JIG == 7):
                $ 1214 "FRM_Reference≔uLM_Cap_SSRack"
                global FRM_Reference=uLM_Cap_SSRack
              end
            end
            $ 1217 "PSE_T≔pose_trans(pose_inv(FRM_Reference), CAM_OBJ_Pose)"
            global PSE_T= pose_trans ( pose_inv (FRM_Reference), CAM_OBJ_Pose)
            $ 1218 "CAM_Result.append(get_pattern_counter(PSE_T, 'X', pattern=[10, 5], patternsize=[0.181, 0.081]))"
            CAM_Result.append(get_pattern_counter(PSE_T, "X", pattern=[10, 5], patternsize=[0.181, 0.081]))
            $ 1219 "PRC_CntDetect≔PRC_CntDetect+1"
            global PRC_CntDetect=PRC_CntDetect+1
          end
          $ 1220 "CAM_Done≔ True "
          global CAM_Done=  True
        else:
          $ 1221 "ElseIf CAM_Captures≥CAM_PRM_Retries"
          if (CAM_Captures >= CAM_PRM_Retries):
            $ 1222 "CAM_Done≔ True "
            global CAM_Done=  True
          else:
            $ 1223 "Else" "noBreak"
            $ 1224 "CAM_Captures≔CAM_Captures+1"
            global CAM_Captures=CAM_Captures+1
          end
        end
      end
    end
    $ 1225 "'=========='"
    # '=========='
    $ 1226 "PostSettings"
    $ 1227 "FRM_Reference≔p[0,0,0,0,0,0]"
    global FRM_Reference=p[0,0,0,0,0,0]
    $ 1228 "Set"
    set_tcp(p[0.0,0.0,0.161,3.1415,0.0,0.0])
    $ 1229 "CAM_Pose≔p[0,0,0,0,0,0]"
    global CAM_Pose=p[0,0,0,0,0,0]
    $ 1230 "Action≔0"
    global Action=0
    $ 1231 "Action_Info≔''"
    global Action_Info=""
  end
  def Sub_AMR_MiR_V3():
    $ 1232 "Sub_AMR_MiR_V3" "noBreak"
    $ 1233 "PreSettings"
    $ 1234 "AMR_TargetList≔[1,2,3,4,5,21,22,23,24,31,32,33,34,35,36,37,38,41]"
    global AMR_TargetList=[1,2,3,4,5,21,22,23,24,31,32,33,34,35,36,37,38,41]
    $ 1235 "AMR_Done≔ False "
    global AMR_Done=  False
    $ 1236 "AMR_PosActual≔T2O_Current_Pos"
    global AMR_PosActual=modbus_get_signal_status("T2O_Current_Pos")
    $ 1237 "AMR_Attemps≔T2O_Nav_Attemps"
    global AMR_Attemps=modbus_get_signal_status("T2O_Nav_Attemps")
    $ 1238 "AMR_Battery≔MiR_Battery_Lvl"
    global AMR_Battery=modbus_get_signal_status("MiR_Battery_Lvl")
    $ 1239 "AMR_Charging≔(T2O_Charging≟1)"
    global AMR_Charging=(modbus_get_signal_status("T2O_Charging") == 1)
    $ 1240 "AMR_Position≔struct(position_identifier=T2O_Current_Pos, x1=MiR_Position_X1, x2=MiR_Position_X2, y1=MiR_Position_Y1, y2=MiR_Position_Y2, theta1=MiR_Theta_1, theta2=MiR_Theta_2) "
    global AMR_Position=struct(position_identifier=modbus_get_signal_status("T2O_Current_Pos"), x1=modbus_get_signal_status("MiR_Position_X1"), x2=modbus_get_signal_status("MiR_Position_X2"), y1=modbus_get_signal_status("MiR_Position_Y1"), y2=modbus_get_signal_status("MiR_Position_Y2"), theta1=modbus_get_signal_status("MiR_Theta_1"), theta2=modbus_get_signal_status("MiR_Theta_2"))
    $ 1241 "If MiR_Mode≠7"
    if (modbus_get_signal_status("MiR_Mode") != 7):
      $ 1242 "Error"
      $ 1243 "set_error(ERROR_AMR_WRONG_MODE)"
      set_error(ERROR_AMR_WRONG_MODE)
      $ 1244 "AMR_Done≔ True "
      global AMR_Done=  True
    end
    $ 1245 "'=========='"
    # '=========='
    $ 1246 "Switch STATE"
    switch_1 = STATE
    $ 1247 "Case 1"
    if (1 == switch_1):
      $ 1248 "stopping"
      $ 1249 "If T2O_Done≟1 and O2T_Acknowledge≟0"
      if (modbus_get_signal_status("T2O_Done") == 1  and  modbus_get_signal_status("O2T_Acknowledge") == 0):
        $ 1250 "Set O2T_Acknowledge=1"
        modbus_set_output_register("O2T_Acknowledge", 1)
      end
      $ 1251 "Set MiR_CMD_Stop=On"
      modbus_set_output_signal("MiR_CMD_Stop", True)
      $ 1252 "AMR_Position.position_identifier = 0"
      AMR_Position.position_identifier = 0
      $ 1253 "AMR_Done≔ True "
      global AMR_Done=  True
    elif (2 == switch_1):
      $ 1254 "Case 2"
      $ 1255 "stopped"
      $ 1256 "If MiR_State≠3 and MiR_State≠5"
      if (modbus_get_signal_status("MiR_State") != 3  and  modbus_get_signal_status("MiR_State") != 5):
        $ 1257 "Set MiR_CMD_Stop=Off"
        modbus_set_output_signal("MiR_CMD_Stop", False)
      end
    elif (3 == switch_1):
      $ 1258 "Case 3"
      $ 1259 "resetting"
      $ 1260 "Set O2T_Mis_Main=Off"
      modbus_set_output_signal("O2T_Mis_Main", False)
      $ 1261 "Set O2T_Mis_Charge=Off"
      modbus_set_output_signal("O2T_Mis_Charge", False)
      $ 1262 "If MiR_Mis_Queue>0"
      if (modbus_get_signal_status("MiR_Mis_Queue")>0):
        $ 1263 "Set MiR_CMD_Clear_Q=On"
        modbus_set_output_signal("MiR_CMD_Clear_Q", True)
        $ 1264 "Wait MiR_Mis_Queue≟0"
        while (not(modbus_get_signal_status("MiR_Mis_Queue") == 0)):
          sync()
        end
        $ 1265 "Set MiR_CMD_Clear_Q=Off"
        modbus_set_output_signal("MiR_CMD_Clear_Q", False)
      end
      $ 1266 "If MiR_Error_ID≠0"
      if (modbus_get_signal_status("MiR_Error_ID") != 0):
        $ 1267 "Set MiR_CMD_Clear_E=On"
        modbus_set_output_signal("MiR_CMD_Clear_E", True)
        $ 1268 "Wait MiR_Error_ID≟0"
        while (not(modbus_get_signal_status("MiR_Error_ID") == 0)):
          sync()
        end
        $ 1269 "Set MiR_CMD_Clear_E=Off"
        modbus_set_output_signal("MiR_CMD_Clear_E", False)
      end
      $ 1270 "Set O2T_Action=0"
      modbus_set_output_register("O2T_Action", 0)
      $ 1271 "Set O2T_Acknowledge=0"
      modbus_set_output_register("O2T_Acknowledge", 0)
      $ 1272 "Set O2T_Target_Pos=0"
      modbus_set_output_register("O2T_Target_Pos", 0)
      $ 1273 "Set O2T_Footprint=0"
      modbus_set_output_register("O2T_Footprint", 0)
      $ 1274 "Set O2T_ProtectOff=0"
      modbus_set_output_register("O2T_ProtectOff", 0)
      $ 1275 "Set O2T_Dock=0"
      modbus_set_output_register("O2T_Dock", 0)
      $ 1276 "AMR_Attemps≔0"
      global AMR_Attemps=0
      $ 1277 "AMR_PosTarget≔0"
      global AMR_PosTarget=0
      $ 1278 "AMR_Step≔0"
      global AMR_Step=0
      $ 1279 "AMR_AtTarget≔ False "
      global AMR_AtTarget=  False
      $ 1280 "If MiR_State≟4 or MiR_State≟3 or MiR_State≟10"
      if (modbus_get_signal_status("MiR_State") == 4  or  modbus_get_signal_status("MiR_State") == 3  or  modbus_get_signal_status("MiR_State") == 10):
        $ 1281 "AMR_Done≔ True "
        global AMR_Done=  True
      end
    elif (5 == switch_1):
      $ 1282 "Case 5"
      $ 1283 "starting"
      $ 1284 "If MiR_State≟4"
      if (modbus_get_signal_status("MiR_State") == 4):
        $ 1285 "Set MiR_CMD_Start=On"
        modbus_set_output_signal("MiR_CMD_Start", True)
        $ 1286 "Wait MiR_State≠4"
        while (not(modbus_get_signal_status("MiR_State") != 4)):
          sync()
        end
        $ 1287 "Set MiR_CMD_Start=Off"
        modbus_set_output_signal("MiR_CMD_Start", False)
        $ 1288 "AMR_Done≔ True "
        global AMR_Done=  True
      else:
        $ 1289 "ElseIf MiR_State≟10"
        if (modbus_get_signal_status("MiR_State") == 10):
          $ 1290 "'MiR in protective stop. Wait'"
          # 'MiR in protective stop. Wait'
          $ 1291 "AMR_Done≔ True "
          global AMR_Done=  True
        else:
          $ 1292 "ElseIf MiR_State≟3"
          if (modbus_get_signal_status("MiR_State") == 3):
            $ 1293 "AMR_Done≔ True "
            global AMR_Done=  True
          end
        end
      end
    elif (6 == switch_1):
      $ 1294 "Case 6"
      $ 1295 "execute"
      $ 1296 "AMR_AtTarget≔(AMR_PosActual≟AMR_PosTarget)"
      global AMR_AtTarget=(AMR_PosActual == AMR_PosTarget)
      $ 1297 "Switch AMR_Step"
      switch_2 = AMR_Step
      $ 1298 "Case 0"
      if (0 == switch_2):
        $ 1299 "If  not AMR_AtTarget"
        if (  not  AMR_AtTarget):
          $ 1300 "AMR_Step≔1"
          global AMR_Step=1
        else:
          $ 1301 "Else" "noBreak"
          $ 1302 "AMR_Done≔ True "
          global AMR_Done=  True
        end
      elif (1 == switch_2):
        $ 1303 "Case 1"
        $ 1304 "general Settings"
        $ 1305 "Set O2T_Acknowledge=0"
        modbus_set_output_register("O2T_Acknowledge", 0)
        $ 1306 "check for error"
        $ 1307 "If OBJ_Picked and MiR_State≟10"
        if (OBJ_Picked  and  modbus_get_signal_status("MiR_State") == 10):
          $ 1308 "Error"
          $ 1309 "set_error(ERROR_ROBOT_ARM_NOT_IN_HOME_POSE)"
          set_error(ERROR_ROBOT_ARM_NOT_IN_HOME_POSE)
          $ 1310 "Action≔0"
          global Action=0
        else:
          $ 1311 "ElseIf  not found_in_list(AMR_PosTarget, AMR_TargetList)"
          if (  not  found_in_list(AMR_PosTarget, AMR_TargetList)):
            $ 1312 "Error"
            $ 1313 "set_error(ERROR_UNKNOWN_POSE)"
            set_error(ERROR_UNKNOWN_POSE)
            $ 1314 "Action≔0"
            global Action=0
          end
        end
        $ 1315 "If MiR_State≟3"
        if (modbus_get_signal_status("MiR_State") == 3):
          $ 1316 "Set MiR_CMD_Start=Off"
          modbus_set_output_signal("MiR_CMD_Start", False)
          $ 1317 "Switch Action"
          switch_3 = Action
          $ 1318 "Case 51"
          if (51 == switch_3):
            $ 1319 "Charge"
            $ 1320 "'trigger the charging mission'"
            # 'trigger the charging mission'
            $ 1321 "'target pos is predefined'"
            # 'target pos is predefined'
            $ 1322 "Set O2T_Footprint=0"
            modbus_set_output_register("O2T_Footprint", 0)
            $ 1323 "Set O2T_Action=1"
            modbus_set_output_register("O2T_Action", 1)
            $ 1324 "If MiR_Mis_Queue≟0"
            if (modbus_get_signal_status("MiR_Mis_Queue") == 0):
              $ 1325 "Set O2T_Mis_Charge=On"
              modbus_set_output_signal("O2T_Mis_Charge", True)
              $ 1326 "Wait MiR_Mis_Queue≥1"
              while (not(modbus_get_signal_status("MiR_Mis_Queue") >= 1)):
                sync()
              end
              $ 1327 "Set O2T_Mis_Charge=Off"
              modbus_set_output_signal("O2T_Mis_Charge", False)
            end
          elif (52 == switch_3):
            $ 1328 "Case 52"
            $ 1329 "Navigate"
            $ 1330 "'trigger the standard missoin'"
            # 'trigger the standard missoin'
            $ 1331 "Set O2T_Footprint=AMR_FootprintID"
            modbus_set_output_register("O2T_Footprint", AMR_FootprintID)
            $ 1332 "Set O2T_Target_Pos=AMR_PosTarget"
            modbus_set_output_register("O2T_Target_Pos", AMR_PosTarget)
            $ 1333 "Set O2T_Action=2"
            modbus_set_output_register("O2T_Action", 2)
            $ 1334 "If MiR_Mis_Queue≟0"
            if (modbus_get_signal_status("MiR_Mis_Queue") == 0):
              $ 1335 "Set O2T_Mis_Main=On"
              modbus_set_output_signal("O2T_Mis_Main", True)
              $ 1336 "Wait MiR_Mis_Queue≥1"
              while (not(modbus_get_signal_status("MiR_Mis_Queue") >= 1)):
                sync()
              end
              $ 1337 "Set O2T_Mis_Main=Off"
              modbus_set_output_signal("O2T_Mis_Main", False)
            end
          end
        else:
          $ 1338 "ElseIf MiR_State≟4"
          if (modbus_get_signal_status("MiR_State") == 4):
            $ 1339 "Set MiR_CMD_Start=On"
            modbus_set_output_signal("MiR_CMD_Start", True)
          else:
            $ 1340 "ElseIf MiR_State≟5"
            if (modbus_get_signal_status("MiR_State") == 5):
              $ 1341 "AMR_Step≔2"
              global AMR_Step=2
            else:
              $ 1342 "ElseIf MiR_State≟10"
              if (modbus_get_signal_status("MiR_State") == 10):
                $ 1343 "'AMR still in safeguard stop'"
                # 'AMR still in safeguard stop'
              end
            end
          end
        end
      elif (2 == switch_2):
        $ 1344 "Case 2"
        $ 1345 "acknowledge handshake"
        $ 1346 "If T2O_Done≟1 and O2T_Acknowledge≟0"
        if (modbus_get_signal_status("T2O_Done") == 1  and  modbus_get_signal_status("O2T_Acknowledge") == 0):
          $ 1347 "Set O2T_Acknowledge=1"
          modbus_set_output_register("O2T_Acknowledge", 1)
        else:
          $ 1348 "ElseIf T2O_Done≟0 and O2T_Acknowledge≟1"
          if (modbus_get_signal_status("T2O_Done") == 0  and  modbus_get_signal_status("O2T_Acknowledge") == 1):
            $ 1349 "Set O2T_Acknowledge=0"
            modbus_set_output_register("O2T_Acknowledge", 0)
            $ 1350 "AMR_AtTarget≔(AMR_PosActual≟AMR_PosTarget)"
            global AMR_AtTarget=(AMR_PosActual == AMR_PosTarget)
            $ 1351 "AMR_Done≔ True "
            global AMR_Done=  True
          end
        end
      end
      $ 1352 "translate errors"
      $ 1353 "If AMR_Done"
      if (AMR_Done):
        $ 1354 "Switch T2O_Error_ID"
        switch_2 = modbus_get_signal_status("T2O_Error_ID")
        $ 1355 "Case 2003"
        if (2003 == switch_2):
          $ 1356 "error"
          $ 1357 "set_error(ERROR_NOT_DOCKED)"
          set_error(ERROR_NOT_DOCKED)
        elif (2007 == switch_2):
          $ 1358 "Case 2007"
          $ 1359 "error"
          $ 1360 "set_error(ERROR_NOT_REACHABLE_TARGET)"
          set_error(ERROR_NOT_REACHABLE_TARGET)
        elif (2008 == switch_2):
          $ 1361 "Case 2008"
          $ 1362 "error"
          $ 1363 "set_error(ERROR_CHARGING_NOT_STARTED)"
          set_error(ERROR_CHARGING_NOT_STARTED)
        end
      end
    elif (7 == switch_1):
      $ 1364 "Case 7"
      $ 1365 "completing"
      $ 1366 "If MiR_Mis_Queue>0"
      if (modbus_get_signal_status("MiR_Mis_Queue")>0):
        $ 1367 "Set MiR_CMD_Abort=On"
        modbus_set_output_signal("MiR_CMD_Abort", True)
        $ 1368 "Wait MiR_Mis_Queue≟0"
        while (not(modbus_get_signal_status("MiR_Mis_Queue") == 0)):
          sync()
        end
        $ 1369 "Set MiR_CMD_Abort=Off"
        modbus_set_output_signal("MiR_CMD_Abort", False)
      end
      $ 1370 "If MiR_State≟3 or MiR_State≟10"
      if (modbus_get_signal_status("MiR_State") == 3  or  modbus_get_signal_status("MiR_State") == 10):
        $ 1371 "AMR_Done≔ True "
        global AMR_Done=  True
      end
    elif (9 == switch_1):
      $ 1372 "Case 9"
      $ 1373 "holding"
      $ 1374 "Set MiR_CMD_Abort=On"
      modbus_set_output_signal("MiR_CMD_Abort", True)
      $ 1375 "If MiR_State≟3 or MiR_State≟10"
      if (modbus_get_signal_status("MiR_State") == 3  or  modbus_get_signal_status("MiR_State") == 10):
        $ 1376 "Set MiR_CMD_Abort=Off"
        modbus_set_output_signal("MiR_CMD_Abort", False)
        $ 1377 "AMR_Done≔ True "
        global AMR_Done=  True
      end
    elif (11 == switch_1):
      $ 1378 "Case 11"
      $ 1379 "unholding"
      $ 1380 "Set MiR_CMD_Start=On"
      modbus_set_output_signal("MiR_CMD_Start", True)
      $ 1381 "If MiR_State≠4"
      if (modbus_get_signal_status("MiR_State") != 4):
        $ 1382 "Set MiR_CMD_Start=Off"
        modbus_set_output_signal("MiR_CMD_Start", False)
        $ 1383 "AMR_Step≔0"
        global AMR_Step=0
        $ 1384 "AMR_Done≔ True "
        global AMR_Done=  True
      end
    elif (12 == switch_1):
      $ 1385 "Case 12"
      $ 1386 "suspending"
      $ 1387 "'none'"
      # 'none'
    elif (14 == switch_1):
      $ 1388 "Case 14"
      $ 1389 "unsuspending"
      $ 1390 "'none'"
      # 'none'
    elif (15 == switch_1):
      $ 1391 "Case 15"
      $ 1392 "aborting"
      $ 1393 "Set MiR_CMD_Abort=On"
      modbus_set_output_signal("MiR_CMD_Abort", True)
      $ 1394 "Wait MiR_State≟3"
      while (not(modbus_get_signal_status("MiR_State") == 3)):
        sync()
      end
      $ 1395 "Set MiR_CMD_Abort=Off"
      modbus_set_output_signal("MiR_CMD_Abort", False)
    elif (17 == switch_1):
      $ 1396 "Case 17"
      $ 1397 "clearing"
      $ 1398 "If MiR_Error_ID≠0"
      if (modbus_get_signal_status("MiR_Error_ID") != 0):
        $ 1399 "Set MiR_CMD_Clear_E=On"
        modbus_set_output_signal("MiR_CMD_Clear_E", True)
        $ 1400 "Wait MiR_Error_ID≟0"
        while (not(modbus_get_signal_status("MiR_Error_ID") == 0)):
          sync()
        end
        $ 1401 "Set MiR_CMD_Clear_E=Off"
        modbus_set_output_signal("MiR_CMD_Clear_E", False)
      end
      $ 1402 "If MiR_Error_ID≟0"
      if (modbus_get_signal_status("MiR_Error_ID") == 0):
        $ 1403 "AMR_Done≔ True "
        global AMR_Done=  True
      end
    end
    $ 1404 "'=========='"
    # '=========='
    $ 1405 "PostSettings"
    $ 1406 "AMR_Position≔struct(position_identifier=T2O_Current_Pos, x1=MiR_Position_X1, x2=MiR_Position_X2, y1=MiR_Position_Y1, y2=MiR_Position_Y2, theta1=MiR_Theta_1, theta2=MiR_Theta_2) "
    global AMR_Position=struct(position_identifier=modbus_get_signal_status("T2O_Current_Pos"), x1=modbus_get_signal_status("MiR_Position_X1"), x2=modbus_get_signal_status("MiR_Position_X2"), y1=modbus_get_signal_status("MiR_Position_Y1"), y2=modbus_get_signal_status("MiR_Position_Y2"), theta1=modbus_get_signal_status("MiR_Theta_1"), theta2=modbus_get_signal_status("MiR_Theta_2"))
  end
  def Sub_Action_V4():
    $ 1407 "Sub_Action_V4" "noBreak"
    $ 1408 "PreSettings"
    $ 1409 "init poses"
    $ 1410 "PSE_A≔p[0,0,0,0,0,0]"
    global PSE_A=p[0,0,0,0,0,0]
    $ 1411 "PSE_A_H≔p[0,0,0,0,0,0]"
    global PSE_A_H=p[0,0,0,0,0,0]
    $ 1412 "PSE_T≔p[0,0,0,0,0,0]"
    global PSE_T=p[0,0,0,0,0,0]
    $ 1413 "PSE_T_H≔p[0,0,0,0,0,0]"
    global PSE_T_H=p[0,0,0,0,0,0]
    $ 1414 "PSE_G≔p[0,0,0,0,0,0]"
    global PSE_G=p[0,0,0,0,0,0]
    $ 1415 "PSE_G_H≔p[0,0,0,0,0,0]"
    global PSE_G_H=p[0,0,0,0,0,0]
    $ 1416 "PSE_R≔p[0,0,0,0,0,0]"
    global PSE_R=p[0,0,0,0,0,0]
    $ 1417 "PSE_R_H≔p[0,0,0,0,0,0]"
    global PSE_R_H=p[0,0,0,0,0,0]
    $ 1418 "JNT_Q≔[0,0,0,0,0,0]"
    global JNT_Q=[0,0,0,0,0,0]
    $ 1419 "JNT_S≔[0,0,0,0,0,0]"
    global JNT_S=[0,0,0,0,0,0]
    $ 1420 "Gripping parameters"
    $ 1421 "OBJ = find_object_by_type(OBJs, OBJ_Type)"
    OBJ = find_object_by_type(OBJs, OBJ_Type)
    $ 1422 "GRP_Open_Pos≔OBJ.dimension.diameter * 1000 + 6"
    global GRP_Open_Pos=OBJ.dimension.diameter * 1000 + 6
    $ 1423 "GRP_Offset≔OBJ.gripper_offset"
    global GRP_Offset=OBJ.gripper_offset
    $ 1424 "rq_set_force_norm(50)"
     rq_set_force_norm (50)
    $ 1425 "rq_set_speed_norm(50)"
     rq_set_speed_norm (50)
    $ 1426 "Switch ITM_ID"
    switch_1 = ITM_ID
    $ 1427 "Case 1"
    if (1 == switch_1):
      $ 1428 "uML"
      $ 1429 "JIG2 = find_object_by_type(JIGs, JIG)"
      JIG2 = find_object_by_type(JIGs, JIG)
      $ 1430 "JIG_Offset≔JIG2.jig_offset"
      global JIG_Offset=JIG2.jig_offset
      $ 1431 "Switch JIG"
      switch_2 = JIG
      $ 1432 "Case 1"
      if (1 == switch_2):
        $ 1433 "3FG"
        $ 1434 "define poses"
        $ 1435 "FRM_Reference≔ULM_3FG"
        global FRM_Reference=ULM_3FG
        $ 1436 "JNT_Q≔JNT_HOME"
        global JNT_Q=JNT_HOME
        $ 1437 "PSE_T≔pose_trans(GRP_Offset, JIG_Offset)"
        global PSE_T= pose_trans (GRP_Offset, JIG_Offset)
        $ 1438 "PSE_A≔pose_trans(PSE_T, p[0,0,0.100,0,0,0])"
        global PSE_A= pose_trans (PSE_T, p[0,0,0.100,0,0,0])
        $ 1439 "PSE_R≔pose_add(PSE_T, p[0,0,0.100,0,0,0])"
        global PSE_R= pose_add (PSE_T, p[0,0,0.100,0,0,0])
      elif (2 == switch_2):
        $ 1440 "Case 2"
        $ 1441 "Input"
        $ 1442 "'CHANGE THE REFERENCE TO THE FRAME TO MOVE IN'"
        # 'CHANGE THE REFERENCE TO THE FRAME TO MOVE IN'
        $ 1443 "define poses"
        $ 1444 "FRM_Reference≔ULM_Input"
        global FRM_Reference=ULM_Input
        $ 1445 "PSE_T≔pose_trans(pose_trans(get_pattern_pos_rectangle(OBJ_Nbr, 'X', [10,5], patternsize=[0.181,0.081]), GRP_Offset), JIG_Offset)"
        global PSE_T= pose_trans ( pose_trans (get_pattern_pos_rectangle(OBJ_Nbr, "X", [10,5], patternsize=[0.181,0.081]), GRP_Offset), JIG_Offset)
        $ 1446 "If Action≟1"
        if (Action == 1):
          $ 1447 "PSE_R≔pose_add(PSE_T, p[0,0,0.200,0,0,0])"
          global PSE_R= pose_add (PSE_T, p[0,0,0.200,0,0,0])
          $ 1448 "PSE_A≔pose_add(PSE_T, p[0,0,0.100,0,0,0])"
          global PSE_A= pose_add (PSE_T, p[0,0,0.100,0,0,0])
        else:
          $ 1449 "ElseIf Action≟2"
          if (Action == 2):
            $ 1450 "PSE_R≔pose_add(PSE_T, p[0,0,0.100,0,0,0])"
            global PSE_R= pose_add (PSE_T, p[0,0,0.100,0,0,0])
            $ 1451 "PSE_A≔pose_add(PSE_T, p[0,0,0.200,0,0,0])"
            global PSE_A= pose_add (PSE_T, p[0,0,0.200,0,0,0])
          end
        end
      elif (3 == switch_2):
        $ 1452 "Case 3"
        $ 1453 "Output"
        $ 1454 "'CHANGE THE REFERENCE TO THE FRAME TO MOVE IN'"
        # 'CHANGE THE REFERENCE TO THE FRAME TO MOVE IN'
        $ 1455 "define poses"
        $ 1456 "FRM_Reference≔ULM_Output"
        global FRM_Reference=ULM_Output
        $ 1457 "PSE_T≔pose_trans(pose_trans(get_pattern_pos_rectangle(OBJ_Nbr, 'X', [10,5], patternsize=[0.181,0.081]), GRP_Offset), JIG_Offset)"
        global PSE_T= pose_trans ( pose_trans (get_pattern_pos_rectangle(OBJ_Nbr, "X", [10,5], patternsize=[0.181,0.081]), GRP_Offset), JIG_Offset)
        $ 1459 "If Action≟1"
        if (Action == 1):
          $ 1460 "PSE_R≔pose_add(PSE_T, p[0,0,0.200,0,0,0])"
          global PSE_R= pose_add (PSE_T, p[0,0,0.200,0,0,0])
          $ 1461 "PSE_A≔pose_add(PSE_T, p[0,0,0.100,0,0,0])"
          global PSE_A= pose_add (PSE_T, p[0,0,0.100,0,0,0])
        else:
          $ 1462 "ElseIf Action≟2"
          if (Action == 2):
            $ 1463 "PSE_R≔pose_add(PSE_T, p[0,0,0.100,0,0,0])"
            global PSE_R= pose_add (PSE_T, p[0,0,0.100,0,0,0])
            $ 1464 "PSE_A≔pose_add(PSE_T, p[0,0,0.200,0,0,0])"
            global PSE_A= pose_add (PSE_T, p[0,0,0.200,0,0,0])
          end
        end
      elif (4 == switch_2):
        $ 1465 "Case 4"
        $ 1466 "jig centrifuge racks"
        $ 1467 "define poses"
        $ 1468 "FRM_Reference≔ULM_Cent_Racks"
        global FRM_Reference=ULM_Cent_Racks
        $ 1469 "PSE_T≔get_pattern_pos_rectangle(JIG_Slot, 'X', [4,1], patternsize=[0.291,0])"
        global PSE_T=get_pattern_pos_rectangle(JIG_Slot, "X", [4,1], patternsize=[0.291,0])
        $ 1470 "If OBJ_Nbr≠0"
        if (OBJ_Nbr != 0):
          $ 1471 "PSE_T≔pose_trans(pose_trans(PSE_T, get_pattern_pos_rectangle(OBJ_Nbr, 'X', [3,3], patternsize=[0.060,0.060])),p[-0.030, -0.030,0,0,0,3.927])"
          global PSE_T= pose_trans ( pose_trans (PSE_T, get_pattern_pos_rectangle(OBJ_Nbr, "X", [3,3], patternsize=[0.060,0.060])),p[-0.030, -0.030,0,0,0,3.927])
        end
        $ 1472 "PSE_T≔pose_trans(PSE_T, GRP_Offset)"
        global PSE_T= pose_trans (PSE_T, GRP_Offset)
        $ 1473 "If Action≟1"
        if (Action == 1):
          $ 1474 "PSE_R≔pose_add(PSE_T, p[0,0,0.200,0,0,0])"
          global PSE_R= pose_add (PSE_T, p[0,0,0.200,0,0,0])
          $ 1475 "PSE_A≔pose_add(PSE_T, p[0,0,0.100,0,0,0])"
          global PSE_A= pose_add (PSE_T, p[0,0,0.100,0,0,0])
        else:
          $ 1476 "ElseIf Action≟2"
          if (Action == 2):
            $ 1477 "PSE_R≔pose_add(PSE_T, p[0,0,0.100,0,0,0])"
            global PSE_R= pose_add (PSE_T, p[0,0,0.100,0,0,0])
            $ 1478 "PSE_A≔pose_add(PSE_T, p[0,0,0.200,0,0,0])"
            global PSE_A= pose_add (PSE_T, p[0,0,0.200,0,0,0])
          end
        end
      elif (6 == switch_2):
        $ 1479 "Case 6"
        $ 1480 "Caps bin"
        $ 1481 "define poses"
        $ 1482 "'Drop cap'"
        # 'Drop cap'
        $ 1483 "FRM_Reference=ULM_Cap_Bin"
        FRM_Reference=ULM_Cap_Bin
        $ 1484 "PSE_T≔pose_RPY2RotVec(p[0,0,0,0,0,0])"
        global PSE_T=pose_RPY2RotVec(p[0,0,0,0,0,0])
        $ 1485 "PSE_T_H≔pose_add(PSE_T, p[0,0,-0.011,0,0,0])"
        global PSE_T_H= pose_add (PSE_T, p[0,0,-0.011,0,0,0])
        $ 1486 "PSE_A≔pose_trans(PSE_T, p[0,0,0.1,0,0,0])"
        global PSE_A= pose_trans (PSE_T, p[0,0,0.1,0,0,0])
        $ 1487 "PSE_R_H≔pose_add(PSE_T, p[0,0,0.100,0,0,0])"
        global PSE_R_H= pose_add (PSE_T, p[0,0,0.100,0,0,0])
        $ 1488 "PSE_R≔pose_add(PSE_T, p[0,0,0.100,0,0,0])"
        global PSE_R= pose_add (PSE_T, p[0,0,0.100,0,0,0])
      elif (7 == switch_2):
        $ 1489 "Case 7"
      elif (8 == switch_2):
        $ 1514 "Case 8"
        $ 1515 "NoK"
        $ 1516 "define poses"
        $ 1517 "'NoK'"
        # 'NoK'
        $ 1518 "FRM_Reference=ULM_NoK"
        FRM_Reference=ULM_NoK
        $ 1519 "PSE_T≔pose_RPY2RotVec(p[0,0,0,0,0,0])"
        global PSE_T=pose_RPY2RotVec(p[0,0,0,0,0,0])
        $ 1520 "PSE_A≔pose_trans(PSE_T, p[0,0,0.1,0,0,0])"
        global PSE_A= pose_trans (PSE_T, p[0,0,0.1,0,0,0])
        $ 1521 "PSE_R≔pose_add(PSE_T, p[0,0,0.100,0,0,0])"
        global PSE_R= pose_add (PSE_T, p[0,0,0.100,0,0,0])
      elif (9 == switch_2):
        $ 1522 "Case 9"
      elif (10 == switch_2):
        $ 1530 "Case 10"
      elif (11 == switch_2):
        $ 1538 "Case 11"
      elif (12 == switch_2):
        $ 1546 "Case 12"
      end
    elif (2 == switch_1):
      $ 1554 "Case 2"
      $ 1555 "Centrifuge"
      $ 1556 "'CHANGE THE REFERENCE TO THE FRAME TO MOVE IN'"
      # 'CHANGE THE REFERENCE TO THE FRAME TO MOVE IN'
      $ 1557 "define poses"
      $ 1558 "FRM_Reference≔FRM_Centrifuge"
      global FRM_Reference=FRM_Centrifuge
      $ 1559 "PSE_T≔GRP_Offset"
      global PSE_T=GRP_Offset
      $ 1560 "If Action≟8"
      if (Action == 8):
        $ 1561 "PSE_R≔pose_add(PSE_T, p[0,0,0.250,0,0,0])"
        global PSE_R= pose_add (PSE_T, p[0,0,0.250,0,0,0])
        $ 1562 "PSE_A≔pose_add(PSE_T, p[0,0,0.150,0,0,0])"
        global PSE_A= pose_add (PSE_T, p[0,0,0.150,0,0,0])
      else:
        $ 1563 "ElseIf Action≟7"
        if (Action == 7):
          $ 1564 "PSE_R≔pose_add(PSE_T, p[0,0,0.150,0,0,0])"
          global PSE_R= pose_add (PSE_T, p[0,0,0.150,0,0,0])
          $ 1565 "PSE_A≔pose_add(PSE_T, p[0,0,0.250,0,0,0])"
          global PSE_A= pose_add (PSE_T, p[0,0,0.250,0,0,0])
        end
      end
    elif (3 == switch_1):
      $ 1566 "Case 3"
      $ 1567 "Output"
      $ 1568 "'CHANGE THE REFERENCE TO THE FRAME TO MOVE IN'"
      # 'CHANGE THE REFERENCE TO THE FRAME TO MOVE IN'
      $ 1569 "define poses"
      $ 1570 "FRM_Reference≔Base_const"
      global FRM_Reference=p[0.0,0.0,0.0,0.0,0.0,0.0]
      $ 1571 "PSE_T≔p[0,0,0,0,0,0]"
      global PSE_T=p[0,0,0,0,0,0]
      $ 1572 "PSE_A≔pose_add(PSE_T, p[0,0,0.150,0,0,0])"
      global PSE_A= pose_add (PSE_T, p[0,0,0.150,0,0,0])
      $ 1573 "PSE_R≔pose_add(PSE_T, p[0,0,0.100,0,0,0])"
      global PSE_R= pose_add (PSE_T, p[0,0,0.100,0,0,0])
    elif (5 == switch_1):
      $ 1574 "Case 5"
      $ 1575 "Sarstedt Pickup Table"
      $ 1576 "'CHANGE THE REFERENCE TO THE FRAME TO MOVE IN'"
      # 'CHANGE THE REFERENCE TO THE FRAME TO MOVE IN'
      $ 1577 "Switch JIG"
      switch_2 = JIG
      $ 1578 "Case 7"
      if (7 == switch_2):
        $ 1591 "Sarstedt"
        $ 1592 "'CHANGE THE REFERENCE TO THE FRAME TO MOVE IN'"
        # 'CHANGE THE REFERENCE TO THE FRAME TO MOVE IN'
        $ 1598 "If TASK.ID≟10"
        if (TASK.ID == 10):
          $ 1599 "Frame & Position Params"
          $ 1600 "FRM_Reference = CAM_LM_SSRack"
          FRM_Reference = CAM_LM_SSRack
          $ 1601 "PSE_T≔uLM_SS_PickPlc"
          global PSE_T=uLM_SS_PickPlc
          $ 1602 "PSE_A≔pose_trans(PSE_T, p[0,0,0.1,0,0,0])"
          global PSE_A= pose_trans (PSE_T, p[0,0,0.1,0,0,0])
          $ 1603 "PSE_R≔pose_add(PSE_T, p[0,0,0.1,0,0,0])"
          global PSE_R= pose_add (PSE_T, p[0,0,0.1,0,0,0])
        end
      end
    elif (13 == switch_1):
      $ 1610 "Case 13"
      $ 1611 "Sarstedt Pickup Table"
      $ 1612 "'CHANGE THE REFERENCE TO THE FRAME TO MOVE IN'"
      # 'CHANGE THE REFERENCE TO THE FRAME TO MOVE IN'
      $ 1613 "Switch JIG"
      switch_2 = JIG
      $ 1614 "Case 7"
      if (7 == switch_2):
        $ 1627 "Bottle"
        $ 1628 "'CHANGE THE REFERENCE TO THE FRAME TO MOVE IN'"
        # 'CHANGE THE REFERENCE TO THE FRAME TO MOVE IN'
        $ 1634 "If TASK.ID≟43"
        if (TASK.ID == 43):
          $ 1635 "Frame & Position Params"
          $ 1637 "PSE_T≔uLM_SS_PickPlc"
          global PSE_T=uLM_SS_PickPlc
          $ 1638 "PSE_A≔pose_trans(PSE_T, p[0,0,0.1,0,0,0])"
          global PSE_A= pose_trans (PSE_T, p[0,0,0.1,0,0,0])
          $ 1639 "PSE_R≔pose_add(PSE_T, p[0,0,0.1,0,0,0])"
          global PSE_R= pose_add (PSE_T, p[0,0,0.1,0,0,0])
        end
      end
    end
    $ 1646 "Additional check"
    $ 1647 "If  not is_reachable(FRM_Reference,[PSE_A,PSE_A_H,PSE_T,PSE_T_H,PSE_R,PSE_R_H])"
    if (  not  is_reachable(FRM_Reference,[PSE_A,PSE_A_H,PSE_T,PSE_T_H,PSE_R,PSE_R_H])):
      $ 1648 "Error"
      $ 1649 "set_error(ERROR_POSE_NOT_REACHABLE)"
      set_error(ERROR_POSE_NOT_REACHABLE)
      $ 1650 "Action≔0"
      global Action=0
    end
    $ 1651 "'=========='"
    # '=========='
    $ 1652 "Switch Action"
    switch_1 = Action
    $ 1653 "Case 1"
    if (1 == switch_1):
      $ 1654 "Pick"
      $ 1655 "Action_Info≔'pick object'"
      global Action_Info="pick object"
      $ 1656 "do_transition(pose_trans(FRM_Reference, PSE_T), keep_rxry=OBJ_Picked)"
      do_transition( pose_trans (FRM_Reference, PSE_T), keep_rxry=OBJ_Picked)
      $ 1657 "EOAT"
      $ 1658 "If  not OBJ_Picked"
      if (  not  OBJ_Picked):
        $ 1659 "rq_move_and_wait_mm(GRP_Open_Pos)"
         rq_move_and_wait_mm (GRP_Open_Pos)
      end
      $ 1660 "If PSE_A_H≠PSE_Z"
      if (PSE_A_H != PSE_Z):
        $ 1661 "If JNT_Q≠JNT_Z"
        if (JNT_Q != JNT_Z):
          $ 1662 "movej(get_inverse_kin(pose_trans(FRM_Reference, PSE_A_H), qnear=JNT_Q), r=0.050)"
          movej(get_inverse_kin( pose_trans (FRM_Reference, PSE_A_H), qnear=JNT_Q), r=0.050)
        else:
          $ 1663 "Else" "noBreak"
          $ 1664 "movej(pose_trans(FRM_Reference, PSE_A_H), r=0.050)"
          movej( pose_trans (FRM_Reference, PSE_A_H), r=0.050)
        end
      end
      $ 1665 "If PSE_A≠PSE_Z"
      if (PSE_A != PSE_Z):
        $ 1666 "If JNT_Q≠JNT_Z"
        if (JNT_Q != JNT_Z):
          $ 1667 "movej(get_inverse_kin(pose_trans(FRM_Reference, PSE_A), qnear=JNT_Q), r=0.020)"
          movej(get_inverse_kin( pose_trans (FRM_Reference, PSE_A), qnear=JNT_Q), r=0.020)
        else:
          $ 1668 "Else" "noBreak"
          $ 1669 "movej(pose_trans(FRM_Reference, PSE_A), r=0.020)"
          movej( pose_trans (FRM_Reference, PSE_A), r=0.020)
        end
      end
      $ 1670 "MoveL"
      $ 1671 "If PSE_T_H≠PSE_Z"
      if (PSE_T_H != PSE_Z):
        $ 1672 "PSE_T_H" "breakAfter"
        movel(pose_trans(FRM_Reference, PSE_T_H), a=0.5, v=0.4, r=0.01)
      end
      $ 1673 "PSE_T" "breakAfter"
      movel(pose_trans(FRM_Reference, PSE_T), a=0.08, v=0.12)
      $ 1674 "EOAT"
      $ 1675 "rq_set_force_norm(50)"
       rq_set_force_norm (50)
      $ 1676 "rq_close_and_wait()"
       rq_close_and_wait ()
      $ 1677 "OBJ_Picked≔rq_is_object_detected()"
      global OBJ_Picked= rq_is_object_detected ()
      $ 1678 "If  not OBJ_Picked"
      if (  not  OBJ_Picked):
        $ 1679 "set_error(ERROR_NO_OBJECT_TO_PICK)"
        set_error(ERROR_NO_OBJECT_TO_PICK)
      end
      $ 1680 "EXTT"
      $ 1681 "Switch JIG"
      switch_2 = JIG
      $ 1682 "Case 1"
      if (1 == switch_2):
        $ 1683 "3FG"
        $ 1684 "If OBJ_Picked"
        if (OBJ_Picked):
          $ 1685 "Set GRP_3F_Open=On"
          set_standard_digital_out(5, True)
        end
      end
      $ 1686 "If PSE_R_H≠PSE_Z"
      if (PSE_R_H != PSE_Z):
        $ 1687 "PSE_R" "breakAfter"
        movel(pose_trans(FRM_Reference, PSE_R), a=0.5, v=0.4, r=0.01)
        $ 1688 "PSE_R_H" "breakAfter"
        movel(pose_trans(FRM_Reference, PSE_R_H), a=0.5, v=0.4)
      else:
        $ 1689 "Else" "noBreak"
        $ 1690 "PSE_R" "breakAfter"
        movel(pose_trans(FRM_Reference, PSE_R), a=0.5, v=0.4)
      end
    elif (2 == switch_1):
      $ 1691 "Case 2"
      $ 1692 "Place"
      $ 1693 "Action_Info≔'place object'"
      global Action_Info="place object"
      $ 1694 "do_transition(pose_trans(FRM_Reference, PSE_T), keep_rxry=OBJ_Picked)"
      do_transition( pose_trans (FRM_Reference, PSE_T), keep_rxry=OBJ_Picked)
      $ 1695 "EXTT"
      $ 1696 "Switch JIG"
      switch_2 = JIG
      $ 1697 "Case 1"
      if (1 == switch_2):
        $ 1698 "3FG"
        $ 1699 "If OBJ_Picked"
        if (OBJ_Picked):
          $ 1700 "Set GRP_3F_Open=On"
          set_standard_digital_out(5, True)
        end
      end
      $ 1701 "If PSE_A_H≠PSE_Z"
      if (PSE_A_H != PSE_Z):
        $ 1702 "If JNT_Q≠JNT_Z"
        if (JNT_Q != JNT_Z):
          $ 1703 "movej(get_inverse_kin(pose_trans(FRM_Reference, PSE_A_H), qnear=JNT_Q), r=0.050)"
          movej(get_inverse_kin( pose_trans (FRM_Reference, PSE_A_H), qnear=JNT_Q), r=0.050)
        else:
          $ 1704 "Else" "noBreak"
          $ 1705 "movej(pose_trans(FRM_Reference, PSE_A_H), r=0.050)"
          movej( pose_trans (FRM_Reference, PSE_A_H), r=0.050)
        end
      end
      $ 1706 "If PSE_A≠PSE_Z"
      if (PSE_A != PSE_Z):
        $ 1707 "If JNT_Q≠JNT_Z"
        if (JNT_Q != JNT_Z):
          $ 1708 "movej(get_inverse_kin(pose_trans(FRM_Reference, PSE_A), qnear=JNT_Q), r=0.020)"
          movej(get_inverse_kin( pose_trans (FRM_Reference, PSE_A), qnear=JNT_Q), r=0.020)
        else:
          $ 1709 "Else" "noBreak"
          $ 1710 "movej(pose_trans(FRM_Reference, PSE_A), r=0.020)"
          movej( pose_trans (FRM_Reference, PSE_A), r=0.020)
        end
      end
      $ 1711 "MoveL"
      $ 1712 "If PSE_T_H≠PSE_Z"
      if (PSE_T_H != PSE_Z):
        $ 1713 "PSE_T_H" "breakAfter"
        movel(pose_trans(FRM_Reference, PSE_T_H), a=0.5, v=0.4, r=0.01)
      end
      $ 1714 "PSE_T" "breakAfter"
      global move_thread_flag_1714=0
      thread move_thread_1714():
        enter_critical
        move_thread_flag_1714 = 1
        movel(pose_trans(FRM_Reference, PSE_T), a=0.05, v=0.09)
        move_thread_flag_1714 = 2
        exit_critical
      end
      move_thread_flag_1714 = 0
      move_thread_han_1714 = run move_thread_1714()
      while (True):
        local targetTcpDirection=get_target_tcp_speed()
        local stepsToRetract=tool_contact(direction=targetTcpDirection)
        if (stepsToRetract > 0):
          kill move_thread_han_1714
          stopl(0.5)
          $ 1715 "Until (tool_contact_detection)"
          break
        end
        sleep(1.0E-10)
        if (move_thread_flag_1714 > 1):
          join move_thread_han_1714
          break
        end
        sync()
      end
      $ 1716 "Force"
      sleep(0.02)
      zero_ftsensor()
      force_mode(FRM_Reference, [1, 1, 1, 0, 0, 0], [0.0, 0.0, 0.0, 0.0, 0.0, 0.0], 2, [0.1, 0.1, 0.01, 0.3490658503988659, 0.3490658503988659, 0.3490658503988659])
      $ 1717 "PSE_T" "noBreak"
      movel(pose_trans(FRM_Reference, PSE_T), a=0.04, v=0.07)
      end_force_mode()
      stopl(5.0)
      $ 1718 "EXTT"
      $ 1719 "Switch JIG"
      switch_2 = JIG
      $ 1720 "Case 1"
      if (1 == switch_2):
        $ 1721 "3FG"
        $ 1722 "If OBJ_Picked"
        if (OBJ_Picked):
          $ 1723 "Set GRP_3F_Open=Off"
          set_standard_digital_out(5, False)
          $ 1724 "Wait: 0.2"
          sleep(0.2)
        end
      end
      $ 1725 "EOAT"
      $ 1726 "rq_move_and_wait_mm(GRP_Open_Pos)"
       rq_move_and_wait_mm (GRP_Open_Pos)
      $ 1727 "OBJ_Picked≔rq_is_object_detected()"
      global OBJ_Picked= rq_is_object_detected ()
      $ 1728 "If PSE_R_H≠PSE_Z"
      if (PSE_R_H != PSE_Z):
        $ 1729 "PSE_R" "breakAfter"
        movel(pose_trans(FRM_Reference, PSE_R), a=0.5, v=0.4, r=0.01)
        $ 1730 "PSE_R_H" "breakAfter"
        movel(pose_trans(FRM_Reference, PSE_R_H), a=0.5, v=0.4)
      else:
        $ 1731 "Else" "noBreak"
        $ 1732 "PSE_R" "breakAfter"
        movel(pose_trans(FRM_Reference, PSE_R), a=0.5, v=0.4)
      end
    elif (3 == switch_1):
      $ 1733 "Case 3"
      $ 1734 "Push"
      $ 1735 "Action_Info≔'push'"
      global Action_Info="push"
    elif (4 == switch_1):
      $ 1736 "Case 4"
      $ 1737 "Pull"
      $ 1738 "Action_Info≔'pull'"
      global Action_Info="pull"
    elif (6 == switch_1):
      $ 1741 "Case 6"
      $ 1742 "Drop the cap"
      $ 1743 "If JNT_A≠[0,0,0,0,0,0]"
      if (JNT_A != [0,0,0,0,0,0]):
        $ 1744 "MoveJ"
        $ 1745 "JNT_A" "breakAfter"
        movej(JNT_A, a=1.3962634015954636, v=1.7453292519943295, r=0.02)
      else:
        $ 1746 "Else" "noBreak"
        $ 1747 "MoveJ"
        $ 1748 "PSE_A" "breakAfter"
        movej(pose_trans(FRM_Reference, PSE_A), a=1.3962634015954636, v=1.7453292519943295, r=0.02)
      end
      $ 1749 "MoveL"
      $ 1750 "PSE_T" "breakAfter"
      movel(pose_trans(FRM_Reference, PSE_T), a=0.05, v=0.09)
      $ 1751 "'ADD OPEN GRIPPER'"
      # 'ADD OPEN GRIPPER'
      # begin: URCap Program Node
      #   Source: Robotiq_Grippers, 3.17.0.105337, Robotiq Inc.
      #   Type: Gripper
      $ 1752 "Gripper Move10mm (1)"
      if not(gripper_connected[0]):
        popup("Gripper 1 must be connected to run this program.", "No connection", False, True, True)
      end
      if not(rq_is_gripper_activated("1")):
        popup("Gripper 1 is not activated. Go to Installation tab > Gripper to activate it and run the program again.", "Not activated", False, True, True)
      end
      rq_set_pos_spd_for(201, 0, 28, "1")
      rq_wait_pos_spe_for_request(201, 0, 28, "1")
      rq_go_to("1")
      rq_wait("1")
      # end: URCap Program Node
      $ 1753 "PSE_T_H" "breakAfter"
      movel(pose_trans(FRM_Reference, PSE_T_H), a=0.05, v=0.09)
      # begin: URCap Program Node
      #   Source: Robotiq_Grippers, 3.17.0.105337, Robotiq Inc.
      #   Type: Gripper
      $ 1754 "Gripper Move40mm (1)"
      if not(gripper_connected[0]):
        popup("Gripper 1 must be connected to run this program.", "No connection", False, True, True)
      end
      if not(rq_is_gripper_activated("1")):
        popup("Gripper 1 is not activated. Go to Installation tab > Gripper to activate it and run the program again.", "Not activated", False, True, True)
      end
      rq_set_pos_spd_for(63, 0, 28, "1")
      rq_wait_pos_spe_for_request(63, 0, 28, "1")
      rq_go_to("1")
      rq_wait("1")
      # end: URCap Program Node
      $ 1755 "PSE_R" "breakAfter"
      movel(pose_trans(FRM_Reference, PSE_R), a=0.5, v=0.4)
    elif (7 == switch_1):
      $ 1756 "Case 7"
      $ 1757 "Load"
      $ 1758 "Action_Info≔'load object'"
      global Action_Info="load object"
      $ 1759 "do_transition(pose_trans(FRM_Reference, PSE_T), keep_rxry=OBJ_Picked)"
      do_transition( pose_trans (FRM_Reference, PSE_T), keep_rxry=OBJ_Picked)
      $ 1760 "If PSE_A_H≠PSE_Z"
      if (PSE_A_H != PSE_Z):
        $ 1761 "If JNT_Q≠JNT_Z"
        if (JNT_Q != JNT_Z):
          $ 1762 "movej(get_inverse_kin(pose_trans(FRM_Reference, PSE_A_H), qnear=JNT_Q), r=0.050)"
          movej(get_inverse_kin( pose_trans (FRM_Reference, PSE_A_H), qnear=JNT_Q), r=0.050)
        else:
          $ 1763 "Else" "noBreak"
          $ 1764 "movej(pose_trans(FRM_Reference, PSE_A_H), r=0.050)"
          movej( pose_trans (FRM_Reference, PSE_A_H), r=0.050)
        end
      end
      $ 1765 "If PSE_A≠PSE_Z"
      if (PSE_A != PSE_Z):
        $ 1766 "If JNT_Q≠JNT_Z"
        if (JNT_Q != JNT_Z):
          $ 1767 "movej(get_inverse_kin(pose_trans(FRM_Reference, PSE_A), qnear=JNT_Q), r=0.020)"
          movej(get_inverse_kin( pose_trans (FRM_Reference, PSE_A), qnear=JNT_Q), r=0.020)
        else:
          $ 1768 "Else" "noBreak"
          $ 1769 "movej(pose_trans(FRM_Reference, PSE_A), r=0.020)"
          movej( pose_trans (FRM_Reference, PSE_A), r=0.020)
        end
      end
      $ 1770 "MoveL"
      $ 1771 "If PSE_T_H≠PSE_Z"
      if (PSE_T_H != PSE_Z):
        $ 1772 "PSE_T_H" "breakAfter"
        movel(pose_trans(FRM_Reference, PSE_T_H), a=0.5, v=0.4, r=0.01)
      end
      $ 1773 "PSE_T" "breakAfter"
      global move_thread_flag_1773=0
      thread move_thread_1773():
        enter_critical
        move_thread_flag_1773 = 1
        movel(pose_trans(FRM_Reference, PSE_T), a=0.05, v=0.09)
        move_thread_flag_1773 = 2
        exit_critical
      end
      move_thread_flag_1773 = 0
      move_thread_han_1773 = run move_thread_1773()
      while (True):
        local targetTcpDirection=get_target_tcp_speed()
        local stepsToRetract=tool_contact(direction=targetTcpDirection)
        if (stepsToRetract > 0):
          kill move_thread_han_1773
          stopl(0.5)
          $ 1774 "Until (tool_contact_detection)"
          break
        end
        sleep(1.0E-10)
        if (move_thread_flag_1773 > 1):
          join move_thread_han_1773
          break
        end
        sync()
      end
      $ 1775 "Force"
      sleep(0.02)
      zero_ftsensor()
      force_mode(FRM_Reference, [0, 1, 1, 0, 0, 1], [0.0, 0.0, 0.0, 0.0, 0.0, 0.0], 2, [0.1, 0.05, 0.02, 0.3490658503988659, 0.3490658503988659, 3.141592653589793])
      $ 1776 "PSE_T" "noBreak"
      movel(pose_trans(FRM_Reference, PSE_T), a=0.04, v=0.07)
      end_force_mode()
      stopl(5.0)
      $ 1777 "EOAT"
      $ 1778 "rq_move_and_wait_mm(GRP_Open_Pos)"
       rq_move_and_wait_mm (GRP_Open_Pos)
      $ 1779 "OBJ_Picked≔rq_is_object_detected()"
      global OBJ_Picked= rq_is_object_detected ()
      $ 1780 "If PSE_R_H≠PSE_Z"
      if (PSE_R_H != PSE_Z):
        $ 1781 "PSE_R" "breakAfter"
        movel(pose_trans(FRM_Reference, PSE_R), a=0.5, v=0.4, r=0.01)
        $ 1782 "PSE_R_H" "breakAfter"
        movel(pose_trans(FRM_Reference, PSE_R_H), a=0.5, v=0.4)
      else:
        $ 1783 "Else" "noBreak"
        $ 1784 "PSE_R" "breakAfter"
        movel(pose_trans(FRM_Reference, PSE_R), a=0.5, v=0.4)
      end
    elif (8 == switch_1):
      $ 1785 "Case 8"
      $ 1786 "Unload"
      $ 1787 "Action_Info≔'pick object'"
      global Action_Info="pick object"
      $ 1788 "do_transition(pose_trans(FRM_Reference, PSE_T), keep_rxry=OBJ_Picked)"
      do_transition( pose_trans (FRM_Reference, PSE_T), keep_rxry=OBJ_Picked)
      $ 1789 "EOAT"
      $ 1790 "If  not OBJ_Picked"
      if (  not  OBJ_Picked):
        $ 1791 "rq_move_and_wait_mm(GRP_Open_Pos)"
         rq_move_and_wait_mm (GRP_Open_Pos)
      end
      $ 1792 "If PSE_A_H≠PSE_Z"
      if (PSE_A_H != PSE_Z):
        $ 1793 "If JNT_Q≠JNT_Z"
        if (JNT_Q != JNT_Z):
          $ 1794 "movej(get_inverse_kin(pose_trans(FRM_Reference, PSE_A_H), qnear=JNT_Q), r=0.050)"
          movej(get_inverse_kin( pose_trans (FRM_Reference, PSE_A_H), qnear=JNT_Q), r=0.050)
        else:
          $ 1795 "Else" "noBreak"
          $ 1796 "movej(pose_trans(FRM_Reference, PSE_A_H), r=0.050)"
          movej( pose_trans (FRM_Reference, PSE_A_H), r=0.050)
        end
      end
      $ 1797 "If PSE_A≠PSE_Z"
      if (PSE_A != PSE_Z):
        $ 1798 "If JNT_Q≠JNT_Z"
        if (JNT_Q != JNT_Z):
          $ 1799 "movej(get_inverse_kin(pose_trans(FRM_Reference, PSE_A), qnear=JNT_Q), r=0.020)"
          movej(get_inverse_kin( pose_trans (FRM_Reference, PSE_A), qnear=JNT_Q), r=0.020)
        else:
          $ 1800 "Else" "noBreak"
          $ 1801 "movej(pose_trans(FRM_Reference, PSE_A), r=0.020)"
          movej( pose_trans (FRM_Reference, PSE_A), r=0.020)
        end
      end
      $ 1802 "MoveL"
      $ 1803 "If PSE_T_H≠PSE_Z"
      if (PSE_T_H != PSE_Z):
        $ 1804 "PSE_T_H" "breakAfter"
        movel(pose_trans(FRM_Reference, PSE_T_H), a=0.5, v=0.4, r=0.01)
      end
      $ 1805 "PSE_T" "breakAfter"
      movel(pose_trans(FRM_Reference, PSE_T), a=0.08, v=0.12)
      $ 1806 "Force"
      sleep(0.02)
      zero_ftsensor()
      force_mode(FRM_Reference, [1, 1, 0, 0, 0, 0], [0.0, 0.0, 0.0, 0.0, 0.0, 0.0], 2, [0.05, 0.05, 0.1, 0.3490658503988659, 0.3490658503988659, 0.3490658503988659])
      $ 1807 "EOAT" "noBreak"
      $ 1808 "rq_set_force_norm(50)" "noBreak"
       rq_set_force_norm (50)
      $ 1809 "rq_close_and_wait()" "noBreak"
       rq_close_and_wait ()
      $ 1810 "OBJ_Picked≔rq_is_object_detected()" "noBreak"
      global OBJ_Picked= rq_is_object_detected ()
      $ 1811 "If  not OBJ_Picked" "noBreak"
      if (  not  OBJ_Picked):
        $ 1812 "set_error(ERROR_NO_OBJECT_TO_PICK)" "noBreak"
        set_error(ERROR_NO_OBJECT_TO_PICK)
      end
      $ 1813 "If PSE_R_H≠PSE_Z" "noBreak"
      if (PSE_R_H != PSE_Z):
        $ 1814 "PSE_R" "noBreak"
        movel(pose_trans(FRM_Reference, PSE_R), a=0.5, v=0.4, r=0.01)
        $ 1815 "PSE_R_H" "noBreak"
        movel(pose_trans(FRM_Reference, PSE_R_H), a=0.5, v=0.4)
      else:
        $ 1816 "Else" "noBreak"
        $ 1817 "PSE_R" "noBreak"
        movel(pose_trans(FRM_Reference, PSE_R), a=0.5, v=0.4)
      end
      end_force_mode()
      stopl(5.0)
    elif (11 == switch_1):
      $ 1818 "Case 11"
    elif (12 == switch_1):
      $ 1855 "Case 12"
      $ 1856 "Decap"
      $ 1857 "Action_Info≔'decapping'"
      global Action_Info="decapping"
      $ 1858 "Set GRP_3F_Enable=On"
      set_standard_digital_out(4, True)
      $ 1859 "Set GRP_3F_Decap=On"
      set_standard_digital_out(3, True)
      $ 1860 "Force"
      sleep(0.02)
      zero_ftsensor()
      force_mode(tool_pose(), [0, 0, 1, 0, 0, 0], [0.0, 0.0, 5.0, 0.0, 0.0, 0.0], 2, [0.1, 0.1, 0.15, 0.3490658503988659, 0.3490658503988659, 0.3490658503988659])
      $ 1861 "check_decapping(offset=0.015, timeout=5, abort=CMD_Hold)" "noBreak"
      check_decapping(offset=0.015, timeout=5, abort=CMD_Hold)
      end_force_mode()
      stopl(5.0)
      $ 1862 "Set GRP_3F_Decap=Off"
      set_standard_digital_out(3, False)
      $ 1863 "Set GRP_3F_Enable=Off"
      set_standard_digital_out(4, False)
      $ 1864 "MoveL"
      $ 1865 "PSE_R" "breakAfter"
      movel(pose_trans(FRM_Reference, PSE_R), a=0.8, v=0.15)
    elif (13 == switch_1):
      $ 1866 "Case 13"
      $ 1867 "TMR_Barcode: Reset"
      TMR_Barcode = 0
      $ 1868 "Read"
      $ 1869 "TMR_Barcode: Start"
      TMR_Barcode_is_counting = True
      $ 1870 "If TMR_Barcode<PRM_TO_Read_BC"
      global thread_flag_1870=0
      thread Thread_if_1870():
        $ 1871 "KeyenceTrigger"
        $ 1872 "Set OClearResult=HI:Pulse 0.2"
        thread SinglePulse4():
          write_output_boolean_register(2, True)
          sleep(0.2)
          write_output_boolean_register(2, False)
        end
        singlePulse4 = run SinglePulse4()
        $ 1873 "Wait: 0.5"
        sleep(0.5)
        $ 1874 "Set OTriggerBarcode=Off"
        write_output_boolean_register(1, False)
        $ 1875 "Wait: 0.5"
        sleep(0.5)
        $ 1876 "Set OTriggerBarcode=On"
        write_output_boolean_register(1, True)
        $ 1877 "Wait: 0.5"
        sleep(0.5)
        $ 1878 "Preorient"
        $ 1879 "TMR_Barcode: Reset"
        TMR_Barcode = 0
        $ 1880 "If ICmdExctd"
        if (read_input_boolean_register(12)):
          $ 1881 "Set GRP_3F_Decap=On"
          set_standard_digital_out(3, True)
          $ 1882 "Set GRP_3F_Enable=On"
          set_standard_digital_out(4, True)
          $ 1883 "Loop ICmdExctd"
          while (read_input_boolean_register(12)):
            $ 1884 "KeyenceTrigger"
            $ 1885 "Set OClearResult=HI:Pulse 0.1"
            thread SinglePulse5():
              write_output_boolean_register(2, True)
              sleep(0.1)
              write_output_boolean_register(2, False)
            end
            singlePulse5 = run SinglePulse5()
            $ 1886 "Wait: 0.3"
            sleep(0.3)
            $ 1887 "Set OTriggerBarcode=Off"
            write_output_boolean_register(1, False)
            $ 1888 "Wait: 0.3"
            sleep(0.3)
            $ 1889 "Set OTriggerBarcode=On"
            write_output_boolean_register(1, True)
            $ 1890 "Wait: 0.1"
            sleep(0.1)
          end
        end
        $ 1891 "If  not ICmdExctd"
        if (  not  read_input_boolean_register(12)):
          $ 1892 "Set GRP_3F_Decap=On"
          set_standard_digital_out(3, True)
          $ 1893 "Set GRP_3F_Enable=On"
          set_standard_digital_out(4, True)
          $ 1894 "Wait ICmdExctd=HI"
          while (read_input_boolean_register(12) == False):
            sync()
          end
        end
        $ 1895 "Set GRP_3F_Decap=Off"
        set_standard_digital_out(3, False)
        $ 1896 "Set GRP_3F_Enable=Off"
        set_standard_digital_out(4, False)
        $ 1897 "OBJ_Brc_OK≔ True "
        global OBJ_Brc_OK=  True
        thread_flag_1870 = 1
      end
      if (TMR_Barcode<PRM_TO_Read_BC):
        global thread_handler_1870=run Thread_if_1870()
        while (thread_flag_1870 == 0):
          if not(TMR_Barcode<PRM_TO_Read_BC):
            kill thread_handler_1870
            thread_flag_1870 = 2
          else:
            sync()
          end
        end
      else:
        thread_flag_1870 = 2
      end
      if (thread_flag_1870 == 2):
        $ 1898 "Else" "noBreak"
        $ 1899 "exeption"
        $ 1900 "error"
        $ 1902 "OBJ_Brc_OK≔ False "
        global OBJ_Brc_OK=  False
      end
      $ 1903 "Set GRP_3F_Decap=Off"
      set_standard_digital_out(3, False)
      $ 1904 "Set GRP_3F_Enable=Off"
      set_standard_digital_out(4, False)
      $ 1905 "Set OTriggerBarcode=Off"
      write_output_boolean_register(1, False)
    elif (15 == switch_1):
      $ 1906 "Case 15"
      $ 1907 "Detect"
      $ 1908 "Action_Info≔'detect'"
      global Action_Info="detect"
    elif (30 == switch_1):
      $ 1909 "Case 30"
      $ 1910 "Shake"
      $ 1911 "Action_Info≔'shake'"
      global Action_Info="shake"
      $ 1912 "do_transition(pose_trans(FRM_Reference, PSE_T), keep_rxry=OBJ_Picked)"
      do_transition( pose_trans (FRM_Reference, PSE_T), keep_rxry=OBJ_Picked)
      $ 1913 "If PSE_A_H≠PSE_Z"
      if (PSE_A_H != PSE_Z):
        $ 1914 "If JNT_Q≠JNT_Z"
        if (JNT_Q != JNT_Z):
          $ 1915 "movej(get_inverse_kin(pose_trans(FRM_Reference, PSE_A_H), qnear=JNT_Q), r=0.050)"
          movej(get_inverse_kin( pose_trans (FRM_Reference, PSE_A_H), qnear=JNT_Q), r=0.050)
        else:
          $ 1916 "Else" "noBreak"
          $ 1917 "movej(pose_trans(FRM_Reference, PSE_A_H), r=0.050)"
          movej( pose_trans (FRM_Reference, PSE_A_H), r=0.050)
        end
      end
      $ 1918 "If PSE_A≠PSE_Z"
      if (PSE_A != PSE_Z):
        $ 1919 "If JNT_Q≠JNT_Z"
        if (JNT_Q != JNT_Z):
          $ 1920 "movej(get_inverse_kin(pose_trans(FRM_Reference, PSE_A), qnear=JNT_Q), r=0.020)"
          movej(get_inverse_kin( pose_trans (FRM_Reference, PSE_A), qnear=JNT_Q), r=0.020)
        else:
          $ 1921 "Else" "noBreak"
          $ 1922 "movej(pose_trans(FRM_Reference, PSE_A), r=0.020)"
          movej( pose_trans (FRM_Reference, PSE_A), r=0.020)
        end
      end
      $ 1923 "MoveL"
      $ 1924 "If PSE_T_H≠PSE_Z"
      if (PSE_T_H != PSE_Z):
        $ 1925 "PSE_T_H" "breakAfter"
        movel(pose_trans(FRM_Reference, PSE_T_H), a=0.5, v=0.4, r=0.01)
      end
      $ 1926 "PSE_T" "breakAfter"
      movel(pose_trans(FRM_Reference, PSE_T), a=0.08, v=0.12)
      $ 1927 "EXTT"
      $ 1928 "Comment"
      # Comment
      $ 1929 "MoveJ"
      $ 1930 "Waypoint_54" "breakAfter"
      movej(get_inverse_kin(Waypoint_54_p, qnear=Waypoint_54_q), a=1.3962634015954636, v=1.0471975511965976)
      $ 1931 "MoveJ"
      $ 1932 "Waypoint_77" "breakAfter"
      movej(get_inverse_kin(Waypoint_77_p, qnear=Waypoint_77_q), a=1.3962634015954636, v=1.0471975511965976)
      $ 1933 "MoveJ"
      $ 1934 "Waypoint_83" "breakAfter"
      movej(get_inverse_kin(Waypoint_83_p, qnear=Waypoint_83_q), a=1.3962634015954636, v=1.0471975511965976)
      $ 1935 "MoveJ"
      $ 1936 "Waypoint_84" "breakAfter"
      movej(get_inverse_kin(Waypoint_84_p, qnear=Waypoint_84_q), a=1.3962634015954636, v=1.0471975511965976)
      $ 1937 "If PSE_R_H≠PSE_Z"
      if (PSE_R_H != PSE_Z):
        $ 1938 "PSE_R" "breakAfter"
        movel(pose_trans(FRM_Reference, PSE_R), a=0.5, v=0.4, r=0.01)
        $ 1939 "PSE_R_H" "breakAfter"
        movel(pose_trans(FRM_Reference, PSE_R_H), a=0.5, v=0.4)
      else:
        $ 1940 "Else" "noBreak"
        $ 1941 "PSE_R" "breakAfter"
        movel(pose_trans(FRM_Reference, PSE_R), a=0.5, v=0.4)
      end
    elif (31 == switch_1):
      $ 1942 "Case 31"
      $ 1943 "Action_Info≔'Pick_Vial'"
      global Action_Info="Pick_Vial"
      $ 1944 "Pick_Vial"
      # begin: URCap Program Node
      #   Source: Robotiq_Grippers, 3.17.0.105337, Robotiq Inc.
      #   Type: Gripper
      $ 1945 "Gripper Open (1)"
      if not(gripper_connected[0]):
        popup("Gripper 1 must be connected to run this program.", "No connection", False, True, True)
      end
      if not(rq_is_gripper_activated("1")):
        popup("Gripper 1 is not activated. Go to Installation tab > Gripper to activate it and run the program again.", "Not activated", False, True, True)
      end
      rq_set_pos_spd_for(0, 82, 71, "1")
      rq_wait_pos_spe_for_request(0, 82, 71, "1")
      rq_go_to("1")
      rq_wait("1")
      # end: URCap Program Node
      $ 1946 "MoveJ"
      $ 1947 "Vial_above_1" "breakAfter"
      movej(get_inverse_kin(Vial_above_1_p, qnear=Vial_above_1_q), a=0.5235987755982988, v=0.4363323129985824, r=0.05)
      $ 1948 "MoveL"
      $ 1949 "Vial_pick_poi_1" "breakAfter"
      movel(Vial_pick_poi_1_p, a=0.5, v=0.1)
      # begin: URCap Program Node
      #   Source: Robotiq_Grippers, 3.17.0.105337, Robotiq Inc.
      #   Type: Gripper
      $ 1950 "Gripper Close (1)"
      if not(gripper_connected[0]):
        popup("Gripper 1 must be connected to run this program.", "No connection", False, True, True)
      end
      if not(rq_is_gripper_activated("1")):
        popup("Gripper 1 is not activated. Go to Installation tab > Gripper to activate it and run the program again.", "Not activated", False, True, True)
      end
      rq_set_pos_spd_for(255, 71, 84, "1")
      rq_wait_pos_spe_for_request(255, 71, 84, "1")
      rq_go_to("1")
      rq_wait("1")
      # end: URCap Program Node
      $ 1951 "MoveL"
      $ 1952 "Waypoint_86" "breakAfter"
      movel(Waypoint_86_p, a=0.5, v=0.1, r=0.05)
      $ 1953 "Home (Safe)"
      movej([-1.2302089344500047, -1.2969853503591224, -1.875639182904262, -1.539621866126728, 1.5731943360401213, -2.80099559440227], a=1.3962634015954636, v=1.0471975511965976)
    elif (32 == switch_1):
      $ 1954 "Case 32"
      $ 1956 "decap_Vial"
      $ 1957 "Set GRP_3F_Open=On"
      set_standard_digital_out(5, True)
      $ 1958 "MoveJ"
      $ 1959 "Waypoint_87" "breakAfter"
      movej(get_inverse_kin(Waypoint_87_p, qnear=Waypoint_87_q), a=0.5235987755982988, v=0.4363323129985824)
      $ 1960 "MoveL"
      $ 1961 "Vial_3FG_plac_1" "breakAfter"
      movel(Vial_3FG_plac_1_p, a=0.5, v=0.1)
      $ 1962 "Set GRP_3F_Open=Off"
      set_standard_digital_out(5, False)
      $ 1963 "Wait: 0.5"
      sleep(0.5)
      $ 1964 "MoveL"
      $ 1965 "Waypoint_88" "breakAfter"
      movel(Waypoint_88_p, a=0.5, v=0.1, r=0.05)
      $ 1966 "MoveJ"
      $ 1967 "cap_dump_1" "breakAfter"
      movej(get_inverse_kin(cap_dump_1_p, qnear=cap_dump_1_q), a=0.5235987755982988, v=0.4363323129985824)
      # begin: URCap Program Node
      #   Source: Robotiq_Grippers, 3.17.0.105337, Robotiq Inc.
      #   Type: Gripper
      $ 1968 "Gripper Open (1)"
      if not(gripper_connected[0]):
        popup("Gripper 1 must be connected to run this program.", "No connection", False, True, True)
      end
      if not(rq_is_gripper_activated("1")):
        popup("Gripper 1 is not activated. Go to Installation tab > Gripper to activate it and run the program again.", "Not activated", False, True, True)
      end
      rq_set_pos_spd_for(0, 255, 255, "1")
      rq_wait_pos_spe_for_request(0, 255, 255, "1")
      rq_go_to("1")
      rq_wait("1")
      # end: URCap Program Node
      $ 1969 "MoveJ"
      $ 1970 "Waypoint_89" "breakAfter"
